// FunctionBlocks/T_SafeMuting
// Model of the TwinSAFE FB MUTING.
// Suppresses the protective device (OSSDIn) while the muting sensors are actuated in the expected order.
// Sequence (sequential inputs, four sensors, forward):
//   M1 on, M2 on, OSSD blocked, M3 on, M1 off, M4 on, M2 off, OSSD clear, M3 off, M4 off
// Sequence (two sensors: parallel inputs, or sequential with MutingIn3/4 unconnected):
//   S1 on, S2 on, OSSD blocked, S1 off, OSSD clear, S2 off
// Any other change of a sensor or the OSSD during a sequence violates it (diagnostic bit 6).
// The Safety Editor refuses an EDM reset time that is not 0 ms, a multiple of 10 ms and at most 60000 ms:
// the model then reports Error with diagnostic bit 15 instead of running (see T_SafeFunctionBlockBase).
{attribute 'reflection'}
FUNCTION_BLOCK T_SafeMuting EXTENDS T_SafeFunctionBlockBase
VAR_INPUT
    MutingEnable : BOOL; // may be a standard PLC signal
    EDM1 : BOOL; // feedback loop of MuteOut
    EDM2 : BOOL; // feedback loop of MuteDelOut
    MutingIn1 : BOOL;
    MutingIn2 : BOOL;
    OSSDIn1 : BOOL; // protective device channel 1 (TRUE = clear)
    OSSDIn2 : BOOL; // protective device channel 2
    MutingIn3 : BOOL;
    MutingIn4 : BOOL;
    Parameters : ST_SafeMutingParameters;
END_VAR
VAR_OUTPUT
    MutingActive : BOOL; // muting lamp
    MuteOut : BOOL;
    MuteDelOut : BOOL;
END_VAR
VAR
    {attribute 'is_connected' := 'MutingEnable'}
    _mutingEnableConnected : BOOL;
    {attribute 'is_connected' := 'EDM1'}
    _eDM1Connected : BOOL;
    {attribute 'is_connected' := 'EDM2'}
    _eDM2Connected : BOOL;
    {attribute 'is_connected' := 'MutingIn1'}
    _mutingIn1Connected : BOOL;
    {attribute 'is_connected' := 'MutingIn2'}
    _mutingIn2Connected : BOOL;
    {attribute 'is_connected' := 'OSSDIn1'}
    _oSSDIn1Connected : BOOL;
    {attribute 'is_connected' := 'OSSDIn2'}
    _oSSDIn2Connected : BOOL;
    {attribute 'is_connected' := 'MutingIn3'}
    _mutingIn3Connected : BOOL;
    {attribute 'is_connected' := 'MutingIn4'}
    _mutingIn4Connected : BOOL;
    _pairs : ARRAY[1..3] OF T_SafeInputPair; // 1: MutingIn1/2, 2: MutingIn3/4, 3: OSSDIn1/2
    _state : E_SafeMutingState := E_SafeMutingState.Stop;
    _prevState : E_SafeMutingState;
    _filterTimers : ARRAY[1..4] OF TON;
    _filtered : ARRAY[1..4] OF BOOL;
    _sensor : ARRAY[1..4] OF BOOL; // actuated sensors after configuration
    _ossdBlocked : BOOL;
    _sensorCount : USINT;
    _seqSensor : ARRAY[1..10] OF USINT; // 0 = OSSD
    _seqLevel : ARRAY[1..10] OF BOOL;
    _seqLength : USINT;
    _seqIndex : USINT; // consumed events
    _expected : ARRAY[0..4] OF BOOL; // expected level of each signal (0 = OSSD blocked)
    _maxTimer : TON;
    _delayTimer : TON;
    _pendingError : BOOL;
    _edmResetTimer1 : TON;
    _edmResetTimer2 : TON;
    _edm1Dropped : BOOL;
    _edm2Dropped : BOOL;
END_VAR

SUPER^();

METHOD PRIVATE Actual : BOOL
VAR_INPUT
    signal : USINT; // 0 = OSSD blocked, 1..4 = sensor actuated
END_VAR
IF signal = 0 THEN
    Actual := _ossdBlocked;
ELSE
    Actual := _sensor[signal];
END_IF
END_METHOD

METHOD PRIVATE AddEvent
VAR_INPUT
    sensor : USINT; // 0 = OSSD
    level : BOOL; // sensor actuated / OSSD blocked
    backwards : BOOL;
END_VAR
IF sensor = 0 AND Parameters.OssdCheckOptional THEN
    RETURN;
END_IF

IF _seqLength >= 10 THEN
    RETURN;
END_IF

_seqLength := _seqLength + 1;

IF sensor > 0 AND backwards THEN
    _seqSensor[_seqLength] := _sensorCount + 1 - sensor;
ELSE
    _seqSensor[_seqLength] := sensor;
END_IF

_seqLevel[_seqLength] := level;
END_METHOD

// Consumes every expected event that has occurred, then checks that no signal deviates
// from the expected pattern. Returns TRUE when the sequence has been violated.
METHOD PRIVATE Advance : BOOL
VAR
    progressed : BOOL;
    next : USINT;
    k : USINT;
END_VAR
REPEAT
    progressed := FALSE;

    IF _seqIndex < _seqLength THEN
        next := _seqIndex + 1;

        IF Actual(_seqSensor[next]) = _seqLevel[next] THEN
            _expected[_seqSensor[next]] := _seqLevel[next];
            _seqIndex                   := next;
            progressed                  := TRUE;
        END_IF
    END_IF
UNTIL NOT progressed
END_REPEAT

FOR k := 0 TO _sensorCount DO
    IF k = 0 AND Parameters.OssdCheckOptional THEN
        CONTINUE;
    END_IF

    IF Actual(k) <> _expected[k] THEN
        Advance := TRUE;
    END_IF
END_FOR
END_METHOD

METHOD PRIVATE AnySensor : BOOL
VAR
    k : USINT;
END_VAR
FOR k := 1 TO _sensorCount DO
    AnySensor := AnySensor OR _sensor[k];
END_FOR
END_METHOD

// Builds the expected event list for the configured sensor arrangement.
METHOD PRIVATE BuildSequence
VAR_INPUT
    backwards : BOOL;
END_VAR
_seqLength := 0;

IF _sensorCount = 4 THEN
    AddEvent(1, TRUE, backwards);
    AddEvent(2, TRUE, backwards);
    AddEvent(0, TRUE, backwards);
    AddEvent(3, TRUE, backwards);
    AddEvent(1, FALSE, backwards);
    AddEvent(4, TRUE, backwards);
    AddEvent(2, FALSE, backwards);
    AddEvent(0, FALSE, backwards);
    AddEvent(3, FALSE, backwards);
    AddEvent(4, FALSE, backwards);
ELSE
    AddEvent(1, TRUE, backwards);
    AddEvent(2, TRUE, backwards);
    AddEvent(0, TRUE, backwards);
    AddEvent(1, FALSE, backwards);
    AddEvent(0, FALSE, backwards);
    AddEvent(2, FALSE, backwards);
END_IF
END_METHOD

// The EDM reset times must be 0 ms or a multiple of 10 ms up to 60000 ms (Safety Editor: "'Reset Time' parameter ... has to be 0 ms or a multiple of 10 ms and maximal 60000 ms").
METHOD PROTECTED ConfigurationOk : BOOL
IF NOT F_SafeResetTimeOk(Parameters.Edm1ResetTime) THEN
    _configurationFault := 'T_SafeMuting: $'Reset Time$' parameter of EDM1 of MUTING has to be 0 ms or a multiple of 10 ms and maximal 60000 ms';
    RETURN;
ELSIF NOT F_SafeResetTimeOk(Parameters.Edm2ResetTime) THEN
    _configurationFault := 'T_SafeMuting: $'Reset Time$' parameter of EDM2 of MUTING has to be 0 ms or a multiple of 10 ms and maximal 60000 ms';
    RETURN;
END_IF

ConfigurationOk := TRUE;
END_METHOD

// Checks the EDM inputs at restart and records diagnostic bits 4/5 on failure.
METHOD PRIVATE EdmInputsOk : BOOL
EdmInputsOk := TRUE;

IF _eDM1Connected AND NOT EDM1 THEN
    SetDiagBit(4);
    EdmInputsOk := FALSE;
END_IF

IF _eDM2Connected AND NOT EDM2 THEN
    SetDiagBit(5);
    EdmInputsOk := FALSE;
END_IF
END_METHOD

// TRUE when every connected EDM input reads 1 (contactors released).
METHOD PRIVATE EdmInputsTrue : BOOL
EdmInputsTrue := (NOT _eDM1Connected OR EDM1) AND (NOT _eDM2Connected OR EDM2);
END_METHOD

// EL6910 extension: after the outputs switch on, each connected EDM input must drop to FALSE
// within its Reset Time. Returns FALSE (and sets diagnostic bits 4/5) on timeout.
METHOD PRIVATE EdmResetOk : BOOL
EdmResetOk := TRUE;

IF _eDM1Connected AND Parameters.Edm1ResetTime > T#0S THEN
    IF NOT EDM1 THEN
        _edm1Dropped := TRUE;
    END_IF

    _edmResetTimer1(IN := NOT _edm1Dropped, PT := Parameters.Edm1ResetTime);

    IF _edmResetTimer1.Q THEN
        SetDiagBit(4);
        EdmResetOk := FALSE;
    END_IF
END_IF

IF _eDM2Connected AND Parameters.Edm2ResetTime > T#0S THEN
    IF NOT EDM2 THEN
        _edm2Dropped := TRUE;
    END_IF

    _edmResetTimer2(IN := NOT _edm2Dropped, PT := Parameters.Edm2ResetTime);

    IF _edmResetTimer2.Q THEN
        SetDiagBit(5);
        EdmResetOk := FALSE;
    END_IF
END_IF
END_METHOD

METHOD PRIVATE IsMuting : BOOL
IsMuting := (TO_BYTE(_state) >= TO_BYTE(E_SafeMutingState.Muting1)) AND (TO_BYTE(_state) <= TO_BYTE(E_SafeMutingState.Muting9));
END_METHOD

PROPERTY MutingState : E_SafeMutingState
GET
MutingState := _state;
END_GET
END_PROPERTY

// State code for the given number of consumed sequence events.
METHOD PRIVATE MutingStateFor : E_SafeMutingState
VAR_INPUT
    consumed : USINT;
END_VAR
CASE consumed OF
    1:
        MutingStateFor := E_SafeMutingState.Muting1;
    2:
        MutingStateFor := E_SafeMutingState.Muting2;
    3:
        MutingStateFor := E_SafeMutingState.Muting3;
    4:
        MutingStateFor := E_SafeMutingState.Muting4;
    5:
        MutingStateFor := E_SafeMutingState.Muting5;
    6:
        MutingStateFor := E_SafeMutingState.Muting6;
    7:
        MutingStateFor := E_SafeMutingState.Muting7;
    8:
        MutingStateFor := E_SafeMutingState.Muting8;
    9:
        MutingStateFor := E_SafeMutingState.Muting9;
ELSE
    MutingStateFor := E_SafeMutingState.Run;
END_CASE
END_METHOD

METHOD PROTECTED Process
VAR
    raw : ARRAY[1..4] OF BOOL;
    i : USINT;
    acknowledge : BOOL;
    discError : BOOL;
    operating : BOOL;
    startFwd : BOOL;
    startBwd : BOOL;
    k : USINT;
    stateBefore : E_SafeMutingState;
    passes : USINT;
END_VAR
// Debounce of the muting inputs
raw[1] := MutingIn1;
raw[2] := MutingIn2;
raw[3] := MutingIn3;
raw[4] := MutingIn4;

FOR i := 1 TO 4 DO
    _filterTimers[i](IN := (raw[i] <> _filtered[i]), PT := Parameters.FilterTime);

    IF _filterTimers[i].Q OR Parameters.FilterTime = T#0S THEN
        _filtered[i] := raw[i];
    END_IF
END_FOR

acknowledge := (_state = E_SafeMutingState.Error) AND _errAck;
_pairs[1](
    In1 := _filtered[1],
    In2 := _filtered[2],
    Active1 := _mutingIn1Connected,
    Active2 := _mutingIn2Connected,
    MakeContact1 := Parameters.MutingIn1MakeContact,
    MakeContact2 := Parameters.MutingIn2MakeContact,
    DiscrepancyTime := Parameters.MutingDiscrepancyTime1,
    Monitor := _fbRun AND NOT Parameters.SequentialInputs,
    SafeInputsAfterDiscError := Parameters.SafeInputsAfterDiscError,
    Acknowledge := acknowledge
);

_pairs[2](
    In1 := _filtered[3],
    In2 := _filtered[4],
    Active1 := _mutingIn3Connected,
    Active2 := _mutingIn4Connected,
    MakeContact1 := Parameters.MutingIn3MakeContact,
    MakeContact2 := Parameters.MutingIn4MakeContact,
    DiscrepancyTime := Parameters.MutingDiscrepancyTime2,
    Monitor := _fbRun AND NOT Parameters.SequentialInputs,
    SafeInputsAfterDiscError := Parameters.SafeInputsAfterDiscError,
    Acknowledge := acknowledge
);

_pairs[3](
    In1 := OSSDIn1,
    In2 := OSSDIn2,
    Active1 := _oSSDIn1Connected,
    Active2 := _oSSDIn2Connected,
    MakeContact1 := Parameters.OSSDIn1MakeContact,
    MakeContact2 := Parameters.OSSDIn2MakeContact,
    DiscrepancyTime := Parameters.OssdDiscrepancyTime,
    Monitor := _fbRun,
    SafeInputsAfterDiscError := Parameters.SafeInputsAfterDiscError,
    Acknowledge := acknowledge
);

IF Parameters.SequentialInputs THEN
    _sensorCount := SEL(_mutingIn3Connected OR _mutingIn4Connected, 2, 4);
    _sensor[1]   := F_SafeInputValue(_mutingIn1Connected, Parameters.MutingIn1MakeContact, _filtered[1]);
    _sensor[2]   := F_SafeInputValue(_mutingIn2Connected, Parameters.MutingIn2MakeContact, _filtered[2]);
    _sensor[3]   := F_SafeInputValue(_mutingIn3Connected, Parameters.MutingIn3MakeContact, _filtered[3]);
    _sensor[4]   := F_SafeInputValue(_mutingIn4Connected, Parameters.MutingIn4MakeContact, _filtered[4]);
ELSE
    _sensorCount := 2;
    _sensor[1]   := _pairs[1].IsActive AND _pairs[1].AllTrue;
    _sensor[2]   := _pairs[2].IsActive AND _pairs[2].AllTrue;
    _sensor[3]   := FALSE;
    _sensor[4]   := FALSE;
END_IF

_ossdBlocked := NOT _pairs[3].AllTrue;

FOR i := 1 TO 3 DO
    discError := discError OR _pairs[i].DiscrepancyError;
END_FOR

IF NOT _fbRun AND _state <> E_SafeMutingState.Error AND _state <> E_SafeMutingState.Reset THEN
    _state := E_SafeMutingState.Stop;
END_IF

operating := (_state = E_SafeMutingState.Safe) OR (_state = E_SafeMutingState.Run) OR IsMuting();

IF discError THEN
    IF operating THEN
        UpdateDiscrepancyDiag();
        _state := E_SafeMutingState.Error;
    ELSIF _state = E_SafeMutingState.DelayOut THEN
        UpdateDiscrepancyDiag();
        _pendingError := TRUE;
    END_IF
END_IF

passes := 0;

REPEAT
    stateBefore := _state;

    CASE _state OF
        E_SafeMutingState.Stop:
            IF StateChanged() THEN
                SetOutputsSafe();
                MutingActive  := FALSE;
                Error         := FALSE;
                Diag          := 0;
                _pendingError := FALSE;
            END_IF

            IF _fbRun THEN
                _state := E_SafeMutingState.Safe;
            END_IF

        E_SafeMutingState.Safe:
            IF StateChanged() THEN
                SetOutputsSafe();
                MutingActive := FALSE;
            END_IF

            IF NOT _ossdBlocked AND EdmInputsTrue() THEN
                _state := E_SafeMutingState.Run;
            END_IF

        E_SafeMutingState.Run:
            IF StateChanged() THEN
                MuteOut      := TRUE;
                MuteDelOut   := TRUE;
                MutingActive := FALSE;
                StartEdmResetMonitoring();
                _seqIndex := 0;
                _maxTimer(IN := FALSE, PT := Parameters.MaxMutingTime);
            END_IF

            startFwd := _sensor[1];
            startBwd := Parameters.BackwardsMode AND _sensor[_sensorCount];

            IF NOT EdmResetOk() THEN
                _state := E_SafeMutingState.Error;
            ELSIF MutingEnable AND (startFwd OR startBwd) THEN
                BuildSequence(startBwd AND NOT startFwd);

                FOR k := 0 TO 4 DO
                    _expected[k] := FALSE;
                END_FOR

                _seqIndex := 0;

                IF Advance() THEN
                    SetDiagBit(6);
                    _state := E_SafeMutingState.Error;
                ELSE
                    _state := MutingStateFor(_seqIndex);
                END_IF
            ELSIF MutingEnable AND AnySensor() THEN
                // a sensor actuated out of order while muting is enabled violates the sequence
                SetDiagBit(6);
                _state := E_SafeMutingState.Error;
            ELSIF _ossdBlocked THEN
                IF Parameters.DelayTime > T#0S THEN
                    _state := E_SafeMutingState.DelayOut;
                ELSE
                    _state := E_SafeMutingState.Safe;
                END_IF
            END_IF

        E_SafeMutingState.Muting1,
        E_SafeMutingState.Muting2,
        E_SafeMutingState.Muting3,
        E_SafeMutingState.Muting4,
        E_SafeMutingState.Muting5,
        E_SafeMutingState.Muting6,
        E_SafeMutingState.Muting7,
        E_SafeMutingState.Muting8,
        E_SafeMutingState.Muting9:
            IF StateChanged() THEN
                MuteOut      := TRUE;
                MuteDelOut   := TRUE;
                MutingActive := TRUE;
            END_IF

            _maxTimer(IN := (Parameters.MaxMutingTime > T#0S), PT := Parameters.MaxMutingTime);

            IF NOT MutingEnable THEN
                // muting withdrawn: the protective device takes over immediately
                IF NOT _ossdBlocked THEN
                    _state := E_SafeMutingState.Run;
                ELSIF Parameters.DelayTime > T#0S THEN
                    _state := E_SafeMutingState.DelayOut;
                ELSE
                    _state := E_SafeMutingState.Safe;
                END_IF
            ELSIF _maxTimer.Q THEN
                SetDiagBit(7);
                _state := E_SafeMutingState.Error;
            ELSIF Advance() THEN
                SetDiagBit(6);
                _state := E_SafeMutingState.Error;
            ELSIF _seqIndex >= _seqLength THEN
                _state := E_SafeMutingState.Run;
            ELSE
                _state := MutingStateFor(_seqIndex);
            END_IF

        E_SafeMutingState.DelayOut:
            IF StateChanged() THEN
                MuteOut      := FALSE;
                MuteDelOut   := TRUE;
                MutingActive := FALSE;
                _delayTimer(IN := FALSE, PT := Parameters.DelayTime);
            END_IF

            _delayTimer(IN := TRUE, PT := Parameters.DelayTime);

            IF _delayTimer.Q THEN
                _state := SEL(_pendingError, E_SafeMutingState.Safe, E_SafeMutingState.Error);
            END_IF

        E_SafeMutingState.Error:
            IF StateChanged() THEN
                SetOutputsSafe();
                MutingActive  := FALSE;
                Error         := TRUE;
                _pendingError := FALSE;
            END_IF

            UpdateDiscrepancyDiag();

            IF _errAck AND NOT discError THEN
                _state := E_SafeMutingState.Reset;
            END_IF

        E_SafeMutingState.Reset:
            IF StateChanged() THEN
                SetOutputsSafe();
                Error := FALSE;
                Diag  := 0;
            END_IF

            IF _errAckFallingEdge THEN
                _state := SEL(_fbRun, E_SafeMutingState.Stop, E_SafeMutingState.Safe);
            END_IF
    END_CASE

    passes := passes + 1;
UNTIL (stateBefore = _state) OR (passes >= 3)
END_REPEAT

State := TO_BYTE(_state);
END_METHOD

METHOD PRIVATE SetOutputsSafe
MuteOut    := FALSE;
MuteDelOut := FALSE;
END_METHOD

METHOD PRIVATE StartEdmResetMonitoring
_edm1Dropped := FALSE;
_edm2Dropped := FALSE;
_edmResetTimer1(IN := FALSE, PT := Parameters.Edm1ResetTime);
_edmResetTimer2(IN := FALSE, PT := Parameters.Edm2ResetTime);
END_METHOD

METHOD PRIVATE StateChanged : BOOL
IF _prevState = _state THEN
    RETURN;
END_IF

_prevState   := _state;
StateChanged := TRUE;
END_METHOD

// Mirrors the discrepancy state of every pair into the diagnostic bits.
METHOD PRIVATE UpdateDiscrepancyDiag
VAR
    i : USINT;
END_VAR
FOR i := 1 TO 3 DO
    IF _pairs[i].DiscrepancyError THEN
        SetDiagBit(SEL(i = 1, SEL(i = 2, 1, 2), 0));

        IF _pairs[i].AwaitingSafeInputs THEN
            SetDiagBit(SEL(i = 1, SEL(i = 2, 9, 10), 8));
        ELSE
            ClearDiagBit(SEL(i = 1, SEL(i = 2, 9, 10), 8));
        END_IF
    END_IF
END_FOR
END_METHOD

END_FUNCTION_BLOCK

// FunctionBlocks/T_SafeOpMode
// Model of the TwinSAFE FB OPMODE (operating mode selector).
// Exactly one connected OpIn input must be TRUE for the matching OpOut to be set.
// Manual restart is active when the Restart port is connected.
// The Safety Editor refuses an OPMODE with fewer than two OpIn ports connected: the model then reports
// Error with diagnostic bit 15 instead of running (see T_SafeFunctionBlockBase).
{attribute 'reflection'}
FUNCTION_BLOCK T_SafeOpMode EXTENDS T_SafeFunctionBlockBase
VAR_INPUT
    Restart : BOOL; // may be a standard PLC signal
    OpIn1 : BOOL;
    OpIn2 : BOOL;
    OpIn3 : BOOL;
    OpIn4 : BOOL;
    OpIn5 : BOOL;
    OpIn6 : BOOL;
    OpIn7 : BOOL;
    OpIn8 : BOOL;
    Parameters : ST_SafeOpModeParameters;
END_VAR
VAR_OUTPUT
    OpOut1 : BOOL;
    OpOut2 : BOOL;
    OpOut3 : BOOL;
    OpOut4 : BOOL;
    OpOut5 : BOOL;
    OpOut6 : BOOL;
    OpOut7 : BOOL;
    OpOut8 : BOOL;
END_VAR
VAR
    {attribute 'is_connected' := 'Restart'}
    _restartConnected : BOOL;
    {attribute 'is_connected' := 'OpIn1'}
    _opIn1Connected : BOOL;
    {attribute 'is_connected' := 'OpIn2'}
    _opIn2Connected : BOOL;
    {attribute 'is_connected' := 'OpIn3'}
    _opIn3Connected : BOOL;
    {attribute 'is_connected' := 'OpIn4'}
    _opIn4Connected : BOOL;
    {attribute 'is_connected' := 'OpIn5'}
    _opIn5Connected : BOOL;
    {attribute 'is_connected' := 'OpIn6'}
    _opIn6Connected : BOOL;
    {attribute 'is_connected' := 'OpIn7'}
    _opIn7Connected : BOOL;
    {attribute 'is_connected' := 'OpIn8'}
    _opIn8Connected : BOOL;
    _state : E_SafeFbState := E_SafeFbState.Stop;
    _prevState : E_SafeFbState;
    _restartPrev : BOOL;
    _discrepancyTimer : TON;
    _modeSelectedBefore : BOOL;
END_VAR

SUPER^();

// At least two OpIn ports must be connected (Safety Editor: "OPMODE does not have at least 2 input ports connected").
METHOD PROTECTED ConfigurationOk : BOOL
VAR
    connectedInputs : USINT;
END_VAR
connectedInputs := BOOL_TO_USINT(_opIn1Connected)
    + BOOL_TO_USINT(_opIn2Connected)
    + BOOL_TO_USINT(_opIn3Connected)
    + BOOL_TO_USINT(_opIn4Connected)
    + BOOL_TO_USINT(_opIn5Connected)
    + BOOL_TO_USINT(_opIn6Connected)
    + BOOL_TO_USINT(_opIn7Connected)
    + BOOL_TO_USINT(_opIn8Connected);

IF connectedInputs < 2 THEN
    _configurationFault := 'T_SafeOpMode: OPMODE does not have at least 2 input ports connected';
    RETURN;
END_IF

ConfigurationOk := TRUE;
END_METHOD

METHOD PROTECTED Process
VAR
    count : USINT;
    selected : USINT;
    exactlyOne : BOOL;
    restartFalling : BOOL;
    monitoring : BOOL;
    operating : BOOL;
    stateBefore : E_SafeFbState;
    passes : USINT;
END_VAR
IF _opIn1Connected AND OpIn1 THEN
    count    := count + 1;
    selected := 1;
END_IF

IF _opIn2Connected AND OpIn2 THEN
    count    := count + 1;
    selected := 2;
END_IF

IF _opIn3Connected AND OpIn3 THEN
    count    := count + 1;
    selected := 3;
END_IF

IF _opIn4Connected AND OpIn4 THEN
    count    := count + 1;
    selected := 4;
END_IF

IF _opIn5Connected AND OpIn5 THEN
    count    := count + 1;
    selected := 5;
END_IF

IF _opIn6Connected AND OpIn6 THEN
    count    := count + 1;
    selected := 6;
END_IF

IF _opIn7Connected AND OpIn7 THEN
    count    := count + 1;
    selected := 7;
END_IF

IF _opIn8Connected AND OpIn8 THEN
    count    := count + 1;
    selected := 8;
END_IF

exactlyOne     := (count = 1);
restartFalling := NOT Restart AND _restartPrev;
_restartPrev   := Restart;

IF NOT _fbRun AND _state <> E_SafeFbState.Error AND _state <> E_SafeFbState.Reset THEN
    _state := E_SafeFbState.Stop;
END_IF

// Discrepancy monitoring of a mode change: none or several inputs set for too long
operating  := (_state = E_SafeFbState.Safe) OR (_state = E_SafeFbState.Start) OR (_state = E_SafeFbState.Run);
monitoring := operating AND _modeSelectedBefore AND NOT exactlyOne AND (Parameters.DiscrepancyTime > T#0S);
_discrepancyTimer(IN := monitoring, PT := Parameters.DiscrepancyTime);

IF _discrepancyTimer.Q AND operating THEN
    SetDiagBit(0);
    _state := E_SafeFbState.Error;
END_IF

passes := 0;

REPEAT
    stateBefore := _state;

    CASE _state OF
        E_SafeFbState.Stop:
            IF StateChanged() THEN
                SetOutputs(0);
                Error               := FALSE;
                Diag                := 0;
                _modeSelectedBefore := FALSE;
            END_IF

            IF _fbRun THEN
                _state := E_SafeFbState.Safe;
            END_IF

        E_SafeFbState.Safe:
            IF StateChanged() THEN
                SetOutputs(0);
            END_IF

            IF exactlyOne THEN
                IF NOT _restartConnected THEN
                    _state := E_SafeFbState.Run;
                ELSIF Restart THEN
                    _state := E_SafeFbState.Start;
                END_IF
            END_IF

        E_SafeFbState.Start:
            IF StateChanged() THEN
                SetOutputs(0);
            END_IF

            IF NOT exactlyOne THEN
                _state := E_SafeFbState.Safe;
            ELSIF restartFalling THEN
                _state := E_SafeFbState.Run;
            END_IF

        E_SafeFbState.Run:
            IF StateChanged() THEN
                _modeSelectedBefore := TRUE;
            END_IF

            IF exactlyOne THEN
                SetOutputs(selected);
            ELSE
                SetOutputs(0);
                _state := E_SafeFbState.Safe;
            END_IF

        E_SafeFbState.Error:
            IF StateChanged() THEN
                SetOutputs(0);
                Error := TRUE;
            END_IF

            IF _errAck THEN
                _state := E_SafeFbState.Reset;
            END_IF

        E_SafeFbState.Reset:
            IF StateChanged() THEN
                Error := FALSE;
                Diag  := 0;
            END_IF

            IF _errAckFallingEdge THEN
                _state := SEL(_fbRun, E_SafeFbState.Stop, E_SafeFbState.Safe);
            END_IF
    END_CASE

    passes := passes + 1;
UNTIL (stateBefore = _state) OR (passes >= 3)
END_REPEAT

State := TO_BYTE(_state);
END_METHOD

METHOD PRIVATE SetOutputs
VAR_INPUT
    selected : USINT; // 0 = all outputs off
END_VAR
OpOut1 := (selected = 1);
OpOut2 := (selected = 2);
OpOut3 := (selected = 3);
OpOut4 := (selected = 4);
OpOut5 := (selected = 5);
OpOut6 := (selected = 6);
OpOut7 := (selected = 7);
OpOut8 := (selected = 8);
END_METHOD

METHOD PRIVATE StateChanged : BOOL
IF _prevState = _state THEN
    RETURN;
END_IF

_prevState   := _state;
StateChanged := TRUE;
END_METHOD

END_FUNCTION_BLOCK

// FunctionBlocks/T_SafeOr
// Model of the TwinSAFE FB OR. Connected inputs are active.
// The Safety Editor refuses an OR with fewer than two OrIn ports connected: the model then reports
// Error with diagnostic bit 15 instead of running (see T_SafeFunctionBlockBase).
{attribute 'reflection'}
FUNCTION_BLOCK T_SafeOr EXTENDS T_SafeFunctionBlockBase
VAR_INPUT
    OrIn1 : BOOL;
    OrIn2 : BOOL;
    OrIn3 : BOOL;
    OrIn4 : BOOL;
    OrIn5 : BOOL;
    OrIn6 : BOOL;
    OrIn7 : BOOL;
    OrIn8 : BOOL;
    Parameters : ST_SafeLogicParameters;
END_VAR
VAR_OUTPUT
    OrOut : BOOL;
END_VAR
VAR
    {attribute 'is_connected' := 'OrIn1'}
    _orIn1Connected : BOOL;
    {attribute 'is_connected' := 'OrIn2'}
    _orIn2Connected : BOOL;
    {attribute 'is_connected' := 'OrIn3'}
    _orIn3Connected : BOOL;
    {attribute 'is_connected' := 'OrIn4'}
    _orIn4Connected : BOOL;
    {attribute 'is_connected' := 'OrIn5'}
    _orIn5Connected : BOOL;
    {attribute 'is_connected' := 'OrIn6'}
    _orIn6Connected : BOOL;
    {attribute 'is_connected' := 'OrIn7'}
    _orIn7Connected : BOOL;
    {attribute 'is_connected' := 'OrIn8'}
    _orIn8Connected : BOOL;
    _state : E_SafeFbState := E_SafeFbState.Stop;
END_VAR

SUPER^();

// At least two OrIn ports must be connected (Safety Editor: "OR does not have at least 2 input ports active and connected").
METHOD PROTECTED ConfigurationOk : BOOL
VAR
    connectedInputs : USINT;
END_VAR
connectedInputs := BOOL_TO_USINT(_orIn1Connected)
    + BOOL_TO_USINT(_orIn2Connected)
    + BOOL_TO_USINT(_orIn3Connected)
    + BOOL_TO_USINT(_orIn4Connected)
    + BOOL_TO_USINT(_orIn5Connected)
    + BOOL_TO_USINT(_orIn6Connected)
    + BOOL_TO_USINT(_orIn7Connected)
    + BOOL_TO_USINT(_orIn8Connected);

IF connectedInputs < 2 THEN
    _configurationFault := 'T_SafeOr: OR does not have at least 2 input ports active and connected';
    RETURN;
END_IF

ConfigurationOk := TRUE;
END_METHOD

METHOD PROTECTED Process
VAR
    result : BOOL;
END_VAR
result := FALSE;
result := result OR F_SafeInputValue(_orIn1Connected, Parameters.In1MakeContact, OrIn1);
result := result OR F_SafeInputValue(_orIn2Connected, Parameters.In2MakeContact, OrIn2);
result := result OR F_SafeInputValue(_orIn3Connected, Parameters.In3MakeContact, OrIn3);
result := result OR F_SafeInputValue(_orIn4Connected, Parameters.In4MakeContact, OrIn4);
result := result OR F_SafeInputValue(_orIn5Connected, Parameters.In5MakeContact, OrIn5);
result := result OR F_SafeInputValue(_orIn6Connected, Parameters.In6MakeContact, OrIn6);
result := result OR F_SafeInputValue(_orIn7Connected, Parameters.In7MakeContact, OrIn7);
result := result OR F_SafeInputValue(_orIn8Connected, Parameters.In8MakeContact, OrIn8);

IF NOT _fbRun THEN
    _state := E_SafeFbState.Stop;
ELSIF result THEN
    _state := E_SafeFbState.Run;
ELSE
    _state := E_SafeFbState.Safe;
END_IF

OrOut := (_state = E_SafeFbState.Run);
Error := FALSE;
Diag  := 0;
State := TO_BYTE(_state);
END_METHOD

END_FUNCTION_BLOCK

// FunctionBlocks/T_SafeSr
// Model of the TwinSAFE FB SR (set dominant latch).
// The Safety Editor refuses an SR with Set or Reset unconnected: the model then reports Error with
// diagnostic bit 15 instead of running (see T_SafeFunctionBlockBase).
{attribute 'reflection'}
FUNCTION_BLOCK T_SafeSr EXTENDS T_SafeFunctionBlockBase
VAR_INPUT
    Set : BOOL;
    Reset : BOOL;
    Parameters : ST_SafeLatchParameters;
END_VAR
VAR_OUTPUT
    SrOut : BOOL;
END_VAR
VAR
    {attribute 'is_connected' := 'Set'}
    _setConnected : BOOL;
    {attribute 'is_connected' := 'Reset'}
    _resetConnected : BOOL;
    _state : E_SafeLatchState := E_SafeLatchState.Stop;
END_VAR

SUPER^();

// Set and Reset must both be connected (Safety Editor: "Inport Set of SR must be connected").
METHOD PROTECTED ConfigurationOk : BOOL
IF NOT _setConnected THEN
    _configurationFault := 'T_SafeSr: Inport Set of SR must be connected';
    RETURN;
ELSIF NOT _resetConnected THEN
    _configurationFault := 'T_SafeSr: Inport Reset of SR must be connected';
    RETURN;
END_IF

ConfigurationOk := TRUE;
END_METHOD

METHOD PROTECTED Process
VAR
    setActive : BOOL;
    resetActive : BOOL;
END_VAR
setActive   := F_SafeInputValue(_setConnected, Parameters.SetMakeContact, Set);
resetActive := F_SafeInputValue(_resetConnected, Parameters.ResetMakeContact, Reset);

IF NOT _fbRun THEN
    _state := E_SafeLatchState.Stop;
ELSE
    IF _state = E_SafeLatchState.Stop THEN
        _state := E_SafeLatchState.Safe;
    END_IF

    IF setActive THEN
        _state := E_SafeLatchState.Set;
    ELSIF resetActive THEN
        _state := E_SafeLatchState.Safe;
    END_IF
END_IF

SrOut := (_state = E_SafeLatchState.Set);
Error := FALSE;
Diag  := 0;
State := TO_BYTE(_state);
END_METHOD

END_FUNCTION_BLOCK

// FunctionBlocks/T_SafeTof
// Model of the TwinSAFE FB TOF (switch-off delay).
// The Safety Editor refuses a TOF with TofIn1 unconnected: the model then reports Error with diagnostic
// bit 15 instead of running (see T_SafeFunctionBlockBase).
{attribute 'reflection'}
FUNCTION_BLOCK T_SafeTof EXTENDS T_SafeFunctionBlockBase
VAR_INPUT
    TofIn1 : BOOL;
    Parameters : ST_SafeTimerParameters;
END_VAR
VAR_OUTPUT
    TofOut : BOOL;
END_VAR
VAR
    {attribute 'is_connected' := 'TofIn1'}
    _tofIn1Connected : BOOL;
    _state : E_SafeFbState := E_SafeFbState.Stop;
    _timer : TOF;
END_VAR

SUPER^();

// TofIn1 must be connected (Safety Editor: "Inport TofIn1 of TOF must be connected").
METHOD PROTECTED ConfigurationOk : BOOL
IF NOT _tofIn1Connected THEN
    _configurationFault := 'T_SafeTof: Inport TofIn1 of TOF must be connected';
    RETURN;
END_IF

ConfigurationOk := TRUE;
END_METHOD

METHOD PROTECTED Process
VAR
    inputActive : BOOL;
END_VAR
inputActive := F_SafeInputValue(_tofIn1Connected, Parameters.MakeContact, TofIn1);

IF NOT _fbRun THEN
    // a stopped FB does not run its delay
    _timer(IN := FALSE, PT := T#0S);
    _state := E_SafeFbState.Stop;
ELSE
    _timer(IN := inputActive, PT := Parameters.DelayTime);

    IF inputActive THEN
        _state := E_SafeFbState.Run;
    ELSIF _timer.Q THEN
        _state := E_SafeFbState.DelayOut;
    ELSE
        _state := E_SafeFbState.Safe;
    END_IF
END_IF

TofOut := (_state = E_SafeFbState.Run) OR (_state = E_SafeFbState.DelayOut);
Error  := FALSE;
Diag   := 0;
State  := TO_BYTE(_state);
END_METHOD

END_FUNCTION_BLOCK

// FunctionBlocks/T_SafeTwoHand
// Model of the TwinSAFE FB TWOHAND (two-hand control).
// Both hands (input pairs) must be actuated, optionally within HandDiscrepancyTime of each other.
// The output can only be set again after both hands were released together.
{attribute 'reflection'}
FUNCTION_BLOCK T_SafeTwoHand EXTENDS T_SafeFunctionBlockBase
VAR_INPUT
    Twohand1 : BOOL; // first hand, channel 1
    Twohand2 : BOOL; // first hand, channel 2
    Twohand3 : BOOL; // second hand, channel 1
    Twohand4 : BOOL; // second hand, channel 2
    Parameters : ST_SafeTwoHandParameters;
END_VAR
VAR_OUTPUT
    TwoHandOut : BOOL;
END_VAR
VAR
    {attribute 'is_connected' := 'Twohand1'}
    _twohand1Connected : BOOL;
    {attribute 'is_connected' := 'Twohand2'}
    _twohand2Connected : BOOL;
    {attribute 'is_connected' := 'Twohand3'}
    _twohand3Connected : BOOL;
    {attribute 'is_connected' := 'Twohand4'}
    _twohand4Connected : BOOL;
    _pairs : ARRAY[1..2] OF T_SafeInputPair;
    _state : E_SafeTwoHandState := E_SafeTwoHandState.Stop;
    _prevState : E_SafeTwoHandState;
    _handTimer : TON;
    _awaitingRelease : BOOL; // between-hands discrepancy error waits for both hands released
END_VAR

SUPER^();

METHOD PROTECTED Process
VAR
    acknowledge : BOOL;
    hand1 : BOOL; // first hand fully actuated
    hand2 : BOOL; // second hand fully actuated
    anyFalse : BOOL; // at least one active input released
    allFalse : BOOL; // every active input released
    discError : BOOL;
    operating : BOOL;
    stateBefore : E_SafeTwoHandState;
    passes : USINT;
END_VAR
acknowledge := (_state = E_SafeTwoHandState.Error) AND _errAck AND NOT _awaitingRelease;
_pairs[1](
    In1 := Twohand1,
    In2 := Twohand2,
    Active1 := _twohand1Connected,
    Active2 := _twohand2Connected,
    MakeContact1 := Parameters.Twohand1MakeContact,
    MakeContact2 := Parameters.Twohand2MakeContact,
    DiscrepancyTime := Parameters.DiscrepancyTime1,
    Monitor := _fbRun,
    SafeInputsAfterDiscError := Parameters.SafeInputsAfterDiscError,
    Acknowledge := acknowledge
);

_pairs[2](
    In1 := Twohand3,
    In2 := Twohand4,
    Active1 := _twohand3Connected,
    Active2 := _twohand4Connected,
    MakeContact1 := Parameters.Twohand3MakeContact,
    MakeContact2 := Parameters.Twohand4MakeContact,
    DiscrepancyTime := Parameters.DiscrepancyTime2,
    Monitor := _fbRun,
    SafeInputsAfterDiscError := Parameters.SafeInputsAfterDiscError,
    Acknowledge := acknowledge
);

hand1     := _pairs[1].IsActive AND _pairs[1].AllTrue;
hand2     := _pairs[2].IsActive AND _pairs[2].AllTrue;
anyFalse  := NOT (_pairs[1].AllTrue AND _pairs[2].AllTrue);
allFalse  := (NOT _pairs[1].IsActive OR _pairs[1].AllFalse) AND (NOT _pairs[2].IsActive OR _pairs[2].AllFalse);
discError := _pairs[1].DiscrepancyError OR _pairs[2].DiscrepancyError;

IF NOT _fbRun AND _state <> E_SafeTwoHandState.Error AND _state <> E_SafeTwoHandState.Reset THEN
    _state := E_SafeTwoHandState.Stop;
END_IF

operating := (_state = E_SafeTwoHandState.Safe)
                 OR (_state = E_SafeTwoHandState.OneButton)
                 OR (_state = E_SafeTwoHandState.TwoButton)
                 OR (_state = E_SafeTwoHandState.Run)
                 OR (_state = E_SafeTwoHandState.Release);

IF discError AND operating THEN
    UpdateDiscrepancyDiag();
    _state := E_SafeTwoHandState.Error;
END_IF

IF _awaitingRelease AND allFalse THEN
    _awaitingRelease := FALSE;
END_IF

passes := 0;

REPEAT
    stateBefore := _state;

    CASE _state OF
        E_SafeTwoHandState.Stop:
            IF StateChanged() THEN
                TwoHandOut := FALSE;
                Error      := FALSE;
                Diag       := 0;
            END_IF

            IF _fbRun THEN
                _state := E_SafeTwoHandState.Safe;
            END_IF

        E_SafeTwoHandState.Safe:
            IF StateChanged() THEN
                TwoHandOut := FALSE;
            END_IF

            IF hand1 THEN
                _state := E_SafeTwoHandState.OneButton;
            ELSIF hand2 THEN
                _state := E_SafeTwoHandState.TwoButton;
            END_IF

        E_SafeTwoHandState.OneButton:
            IF StateChanged() THEN
                _handTimer(IN := FALSE, PT := Parameters.HandDiscrepancyTime);
            END_IF

            _handTimer(IN := (Parameters.HandDiscrepancyTime > T#0S), PT := Parameters.HandDiscrepancyTime);

            IF _handTimer.Q THEN
                SetHandDiscrepancyError();
            ELSIF hand1 AND hand2 THEN
                _state := E_SafeTwoHandState.Run;
            ELSIF hand2 THEN
                // second hand actuated while the first is no longer detected
                SetDiagBit(6);
                _state := E_SafeTwoHandState.Error;
            ELSIF NOT hand1 THEN
                _state := SEL(allFalse, E_SafeTwoHandState.Release, E_SafeTwoHandState.Safe);
            END_IF

        E_SafeTwoHandState.TwoButton:
            IF StateChanged() THEN
                _handTimer(IN := FALSE, PT := Parameters.HandDiscrepancyTime);
            END_IF

            _handTimer(IN := (Parameters.HandDiscrepancyTime > T#0S), PT := Parameters.HandDiscrepancyTime);

            IF _handTimer.Q THEN
                SetHandDiscrepancyError();
            ELSIF hand1 AND hand2 THEN
                _state := E_SafeTwoHandState.Run;
            ELSIF hand1 THEN
                SetDiagBit(6);
                _state := E_SafeTwoHandState.Error;
            ELSIF NOT hand2 THEN
                _state := SEL(allFalse, E_SafeTwoHandState.Release, E_SafeTwoHandState.Safe);
            END_IF

        E_SafeTwoHandState.Run:
            IF StateChanged() THEN
                TwoHandOut := TRUE;
            END_IF

            IF anyFalse THEN
                _state := E_SafeTwoHandState.Release;
            END_IF

        E_SafeTwoHandState.Release:
            IF StateChanged() THEN
                TwoHandOut := FALSE;
            END_IF

            IF allFalse THEN
                _state := E_SafeTwoHandState.Safe;
            END_IF

        E_SafeTwoHandState.Error:
            IF StateChanged() THEN
                TwoHandOut := FALSE;
                Error      := TRUE;
            END_IF

            UpdateDiscrepancyDiag();

            IF _awaitingRelease THEN
                SetDiagBit(10);
            ELSE
                ClearDiagBit(10);
            END_IF

            IF _errAck AND NOT _awaitingRelease AND NOT discError THEN
                _state := E_SafeTwoHandState.Reset;
            END_IF

        E_SafeTwoHandState.Reset:
            IF StateChanged() THEN
                TwoHandOut := FALSE;
                Error      := FALSE;
                Diag       := 0;
            END_IF

            IF _errAckFallingEdge THEN
                _state := SEL(_fbRun, E_SafeTwoHandState.Stop, E_SafeTwoHandState.Safe);
            END_IF
    END_CASE

    passes := passes + 1;
UNTIL (stateBefore = _state) OR (passes >= 3)
END_REPEAT

State := TO_BYTE(_state);
END_METHOD

METHOD PRIVATE SetHandDiscrepancyError
SetDiagBit(2);
_awaitingRelease := Parameters.SafeInputsAfterDiscError;
_state           := E_SafeTwoHandState.Error;
END_METHOD

METHOD PRIVATE StateChanged : BOOL
IF _prevState = _state THEN
    RETURN;
END_IF

_prevState   := _state;
StateChanged := TRUE;
END_METHOD

PROPERTY TwoHandState : E_SafeTwoHandState
GET
TwoHandState := _state;
END_GET
END_PROPERTY

// Mirrors the discrepancy state of every pair into the diagnostic bits.
METHOD PRIVATE UpdateDiscrepancyDiag
VAR
    i : USINT;
END_VAR
FOR i := 1 TO 2 DO
    IF _pairs[i].DiscrepancyError THEN
        SetDiagBit(i - 1);

        IF _pairs[i].AwaitingSafeInputs THEN
            SetDiagBit(i + 7);
        ELSE
            ClearDiagBit(i + 7);
        END_IF
    END_IF
END_FOR
END_METHOD

END_FUNCTION_BLOCK

// FunctionBlocks/T_SafeXor
// Model of the TwinSAFE FB XOR: eight independent exclusive-or pairs. A pair is active when connected.
{attribute 'reflection'}
FUNCTION_BLOCK T_SafeXor EXTENDS T_SafeFunctionBlockBase
VAR_INPUT
    Xor1In1 : BOOL;
    Xor2In1 : BOOL;
    Xor1In2 : BOOL;
    Xor2In2 : BOOL;
    Xor1In3 : BOOL;
    Xor2In3 : BOOL;
    Xor1In4 : BOOL;
    Xor2In4 : BOOL;
    Xor1In5 : BOOL;
    Xor2In5 : BOOL;
    Xor1In6 : BOOL;
    Xor2In6 : BOOL;
    Xor1In7 : BOOL;
    Xor2In7 : BOOL;
    Xor1In8 : BOOL;
    Xor2In8 : BOOL;
END_VAR
VAR_OUTPUT
    XorOut1 : BOOL;
    XorOut2 : BOOL;
    XorOut3 : BOOL;
    XorOut4 : BOOL;
    XorOut5 : BOOL;
    XorOut6 : BOOL;
    XorOut7 : BOOL;
    XorOut8 : BOOL;
END_VAR
VAR
    {attribute 'is_connected' := 'Xor1In1'}
    _xor1In1Connected : BOOL;
    {attribute 'is_connected' := 'Xor1In2'}
    _xor1In2Connected : BOOL;
    {attribute 'is_connected' := 'Xor1In3'}
    _xor1In3Connected : BOOL;
    {attribute 'is_connected' := 'Xor1In4'}
    _xor1In4Connected : BOOL;
    {attribute 'is_connected' := 'Xor1In5'}
    _xor1In5Connected : BOOL;
    {attribute 'is_connected' := 'Xor1In6'}
    _xor1In6Connected : BOOL;
    {attribute 'is_connected' := 'Xor1In7'}
    _xor1In7Connected : BOOL;
    {attribute 'is_connected' := 'Xor1In8'}
    _xor1In8Connected : BOOL;
    {attribute 'is_connected' := 'Xor2In1'}
    _xor2In1Connected : BOOL;
    {attribute 'is_connected' := 'Xor2In2'}
    _xor2In2Connected : BOOL;
    {attribute 'is_connected' := 'Xor2In3'}
    _xor2In3Connected : BOOL;
    {attribute 'is_connected' := 'Xor2In4'}
    _xor2In4Connected : BOOL;
    {attribute 'is_connected' := 'Xor2In5'}
    _xor2In5Connected : BOOL;
    {attribute 'is_connected' := 'Xor2In6'}
    _xor2In6Connected : BOOL;
    {attribute 'is_connected' := 'Xor2In7'}
    _xor2In7Connected : BOOL;
    {attribute 'is_connected' := 'Xor2In8'}
    _xor2In8Connected : BOOL;
    _state : E_SafeFbState := E_SafeFbState.Stop;
END_VAR

SUPER^();

METHOD PROTECTED Process
VAR
    run : BOOL;
END_VAR
run     := _fbRun;
_state  := SEL(run, E_SafeFbState.Stop, E_SafeFbState.Run);
XorOut1 := run AND (_xor1In1Connected OR _xor2In1Connected) AND (Xor1In1 XOR Xor2In1);
XorOut2 := run AND (_xor1In2Connected OR _xor2In2Connected) AND (Xor1In2 XOR Xor2In2);
XorOut3 := run AND (_xor1In3Connected OR _xor2In3Connected) AND (Xor1In3 XOR Xor2In3);
XorOut4 := run AND (_xor1In4Connected OR _xor2In4Connected) AND (Xor1In4 XOR Xor2In4);
XorOut5 := run AND (_xor1In5Connected OR _xor2In5Connected) AND (Xor1In5 XOR Xor2In5);
XorOut6 := run AND (_xor1In6Connected OR _xor2In6Connected) AND (Xor1In6 XOR Xor2In6);
XorOut7 := run AND (_xor1In7Connected OR _xor2In7Connected) AND (Xor1In7 XOR Xor2In7);
XorOut8 := run AND (_xor1In8Connected OR _xor2In8Connected) AND (Xor1In8 XOR Xor2In8);
Error   := FALSE;
Diag    := 0;
State   := TO_BYTE(_state);
END_METHOD

END_FUNCTION_BLOCK

// Project Information/F_GetCompany
// This function has been automatically generated from the project information.
{attribute 'signature_flag' := '1073741824'}
{attribute 'TcGenerated'}
{attribute 'no-analysis'}
FUNCTION F_GetCompany : WSTRING
VAR_INPUT
	
END_VAR

F_GetCompany := "Intecre Ltd";

END_FUNCTION

// Project Information/F_GetTitle
// This function has been automatically generated from the project information.
{attribute 'signature_flag' := '1073741824'}
{attribute 'TcGenerated'}
{attribute 'no-analysis'}
FUNCTION F_GetTitle : WSTRING
VAR_INPUT
	
END_VAR

F_GetTitle := "Intecre.TwinSAFE.Models";

END_FUNCTION

// Project Information/F_GetVersion
// This function has been automatically generated from the project information.
{attribute 'signature_flag' := '1073741824'}
{attribute 'TcGenerated'}
{attribute 'no-analysis'}
FUNCTION F_GetVersion : ST_LibVersion
VAR_INPUT
	
END_VAR

F_GetVersion.iMajor := 0;
F_GetVersion.iMinor := 5;
F_GetVersion.iBuild := 0;
F_GetVersion.iRevision := 3;
F_GetVersion.sVersion := '0.5.0.3';
F_GetVersion.nFlags := 0;

END_FUNCTION

// Tests/User_FB_Tests/T_SafePulse_UserFB_Tests
// Tests of the example user FB T_SafePulse_UserFB: TonOut is a pulse of DelayTime while TonIn1 is held.
FUNCTION_BLOCK T_SafePulse_UserFB_Tests EXTENDS TcUnit.FB_TestSuite
VAR
    // Test_PulseForDelayTimeWhileInputHeld
    group_1 : T_SafeGroup;
    fb_1 : T_SafePulse_UserFB(group := group_1) := (Parameters := (DelayTime := T#100MS));
    state_1 : INT := 10;
    waitTimer_1 : TON;
    // Test_PulseEndsWhenInputDrops
    group_2 : T_SafeGroup;
    fb_2 : T_SafePulse_UserFB(group := group_2) := (Parameters := (DelayTime := T#100MS));
    // Test_StoppedGivesNoOutput
    group_3 : T_SafeGroup;
    fb_3 : T_SafePulse_UserFB(group := group_3) := (Parameters := (DelayTime := T#100MS));
    // Test_InnerBlocksJoinTheGroup
    group_4 : T_SafeGroup;
    fb_4 : T_SafePulse_UserFB(group := group_4);
END_VAR

Test_PulseForDelayTimeWhileInputHeld();
Test_PulseEndsWhenInputDrops();
Test_StoppedGivesNoOutput();
Test_InnerBlocksJoinTheGroup();

METHOD PRIVATE Test_InnerBlocksJoinTheGroup
TcUnit.TEST(__POUNAME());
// assert: the composite registered itself and passed the group on to its TON and AND
AssertEquals_UINT(Expected := 3, Actual := group_4.FunctionBlockCount, Message := 'composite and its two inner blocks registered');
TEST_FINISHED_NAMED(__POUNAME());
END_METHOD

METHOD PRIVATE Test_PulseEndsWhenInputDrops
TcUnit.TEST(__POUNAME());
// act / assert
group_2(Run := TRUE);
fb_2(TonIn1 := TRUE);
AssertEquals_BOOL(Expected := TRUE, Actual := fb_2.TonOut, Message := 'pulse on');
AssertEquals_BOOL(Expected := TRUE, Actual := fb_2.IsRunning, Message := 'reports Run to the group while it runs');
fb_2(TonIn1 := FALSE);
AssertEquals_BOOL(Expected := FALSE, Actual := fb_2.TonOut, Message := 'pulse cut off when the input drops');
TEST_FINISHED_NAMED(__POUNAME());
END_METHOD

METHOD PRIVATE Test_PulseForDelayTimeWhileInputHeld
TcUnit.TEST(__POUNAME());
waitTimer_1();

CASE state_1 OF
    10:
        // act: input on, the pulse starts
        group_1(Run := TRUE);
        fb_1(TonIn1 := TRUE);
        // assert
        AssertEquals_BOOL(Expected := TRUE, Actual := fb_1.TonOut, Message := 'pulse starts with the input');
        state_1 := 20;
        waitTimer_1(IN := TRUE, PT := T#50MS);
    20:
        group_1(Run := TRUE);
        fb_1(TonIn1 := TRUE);

        IF NOT waitTimer_1.Q THEN
            RETURN;
        END_IF

        waitTimer_1(IN := FALSE);
        // assert: still inside the delay time
        AssertEquals_BOOL(Expected := TRUE, Actual := fb_1.TonOut, Message := 'pulse still on inside the delay time');
        state_1 := 30;
        waitTimer_1(IN := TRUE, PT := T#200MS);
    30:
        group_1(Run := TRUE);
        fb_1(TonIn1 := TRUE);

        IF NOT waitTimer_1.Q THEN
            RETURN;
        END_IF

        waitTimer_1(IN := FALSE);
        // assert: the delay has elapsed, the pulse is over although the input is still held
        AssertEquals_BOOL(Expected := FALSE, Actual := fb_1.TonOut, Message := 'pulse ends after the delay time');
        // act: release and re-apply the input
        fb_1(TonIn1 := FALSE);
        AssertEquals_BOOL(Expected := FALSE, Actual := fb_1.TonOut, Message := 'no output with the input off');
        fb_1(TonIn1 := TRUE);
        AssertEquals_BOOL(Expected := TRUE, Actual := fb_1.TonOut, Message := 'a new pulse starts on the next rising edge');
        TEST_FINISHED_NAMED(__POUNAME());
        state_1 := 10;
END_CASE
END_METHOD

METHOD PRIVATE Test_StoppedGivesNoOutput
TcUnit.TEST(__POUNAME());
// act
group_3(Run := FALSE);
fb_3(TonIn1 := TRUE);
// assert
AssertEquals_BOOL(Expected := FALSE, Actual := fb_3.TonOut, Message := 'no output while the group is stopped');
AssertEquals_BOOL(Expected := FALSE, Actual := fb_3.IsRunning, Message := 'not running while the group is stopped');
TEST_FINISHED_NAMED(__POUNAME());
END_METHOD

END_FUNCTION_BLOCK

// Tests/User_FB_Tests/T_SafePulse_UserFB_Tests_CFC
    // CFC twin of T_SafePulse_UserFB_Tests: the same tests drawn as CFC diagrams, the way a TwinSAFE project is authored.
    FUNCTION_BLOCK T_SafePulse_UserFB_Tests_CFC EXTENDS T_SafeCfcTestSuite
    VAR
    // Test_PulseForDelayTimeWhileInputHeld
    group_1 : T_SafeGroup;
    fb_1 : T_SafePulse_UserFB(group := group_1) := (Parameters := (DelayTime := T#100MS));
    trigStart_1 : R_TRIG;
    t1_1 : TON;
    t2_1 : TON;
    trig1_1 : R_TRIG;
    trig2_1 : R_TRIG;
    // Test_PulseEndsWhenInputDrops
    group_2 : T_SafeGroup;
    fb_2 : T_SafePulse_UserFB(group := group_2) := (Parameters := (DelayTime := T#100MS));
    // Test_StoppedGivesNoOutput
    group_3 : T_SafeGroup;
    fb_3 : T_SafePulse_UserFB(group := group_3) := (Parameters := (DelayTime := T#100MS));
    // Test_InnerBlocksJoinTheGroup
    group_4 : T_SafeGroup;
    fb_4 : T_SafePulse_UserFB(group := group_4);
END_VAR

Test_PulseForDelayTimeWhileInputHeld();
Test_PulseEndsWhenInputDrops();
Test_StoppedGivesNoOutput();
Test_InnerBlocksJoinTheGroup();

METHOD PRIVATE Test_InnerBlocksJoinTheGroup
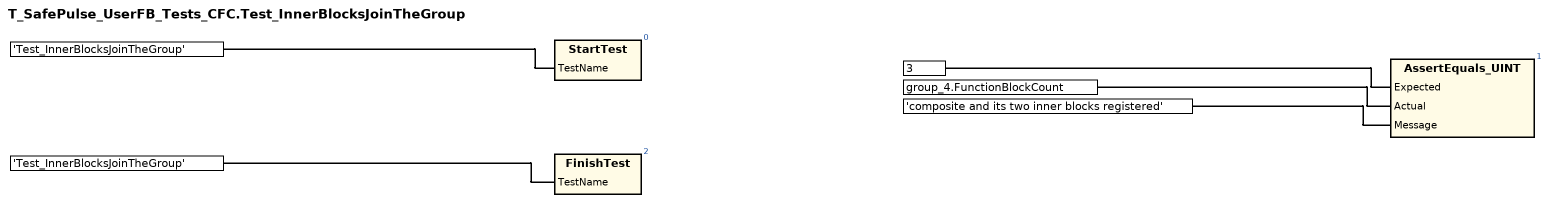
StartTest(TestName := 'Test_InnerBlocksJoinTheGroup');
AssertEquals_UINT(Expected := 3, Actual := group_4.FunctionBlockCount, Message := 'composite and its two inner blocks registered');
FinishTest(TestName := 'Test_InnerBlocksJoinTheGroup');
END_METHOD

METHOD PRIVATE Test_PulseEndsWhenInputDrops
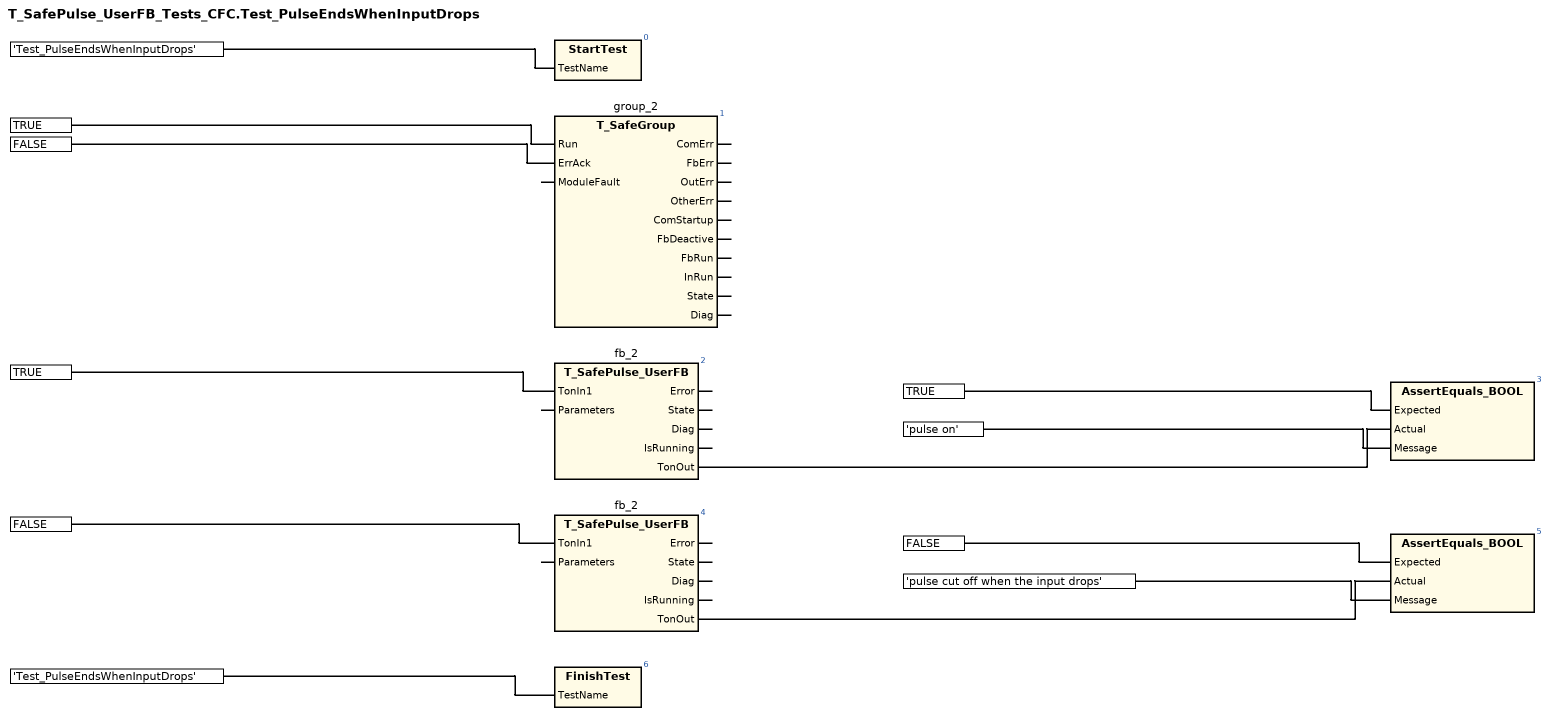
StartTest(TestName := 'Test_PulseEndsWhenInputDrops');
group_2(Run := TRUE, ErrAck := FALSE); // T_SafeGroup
fb_2(TonIn1 := TRUE); // T_SafePulse_UserFB
AssertEquals_BOOL(Expected := TRUE, Actual := fb_2.TonOut, Message := 'pulse on');
fb_2(TonIn1 := FALSE); // T_SafePulse_UserFB
AssertEquals_BOOL(Expected := FALSE, Actual := fb_2.TonOut, Message := 'pulse cut off when the input drops');
FinishTest(TestName := 'Test_PulseEndsWhenInputDrops');
END_METHOD

METHOD PRIVATE Test_PulseForDelayTimeWhileInputHeld
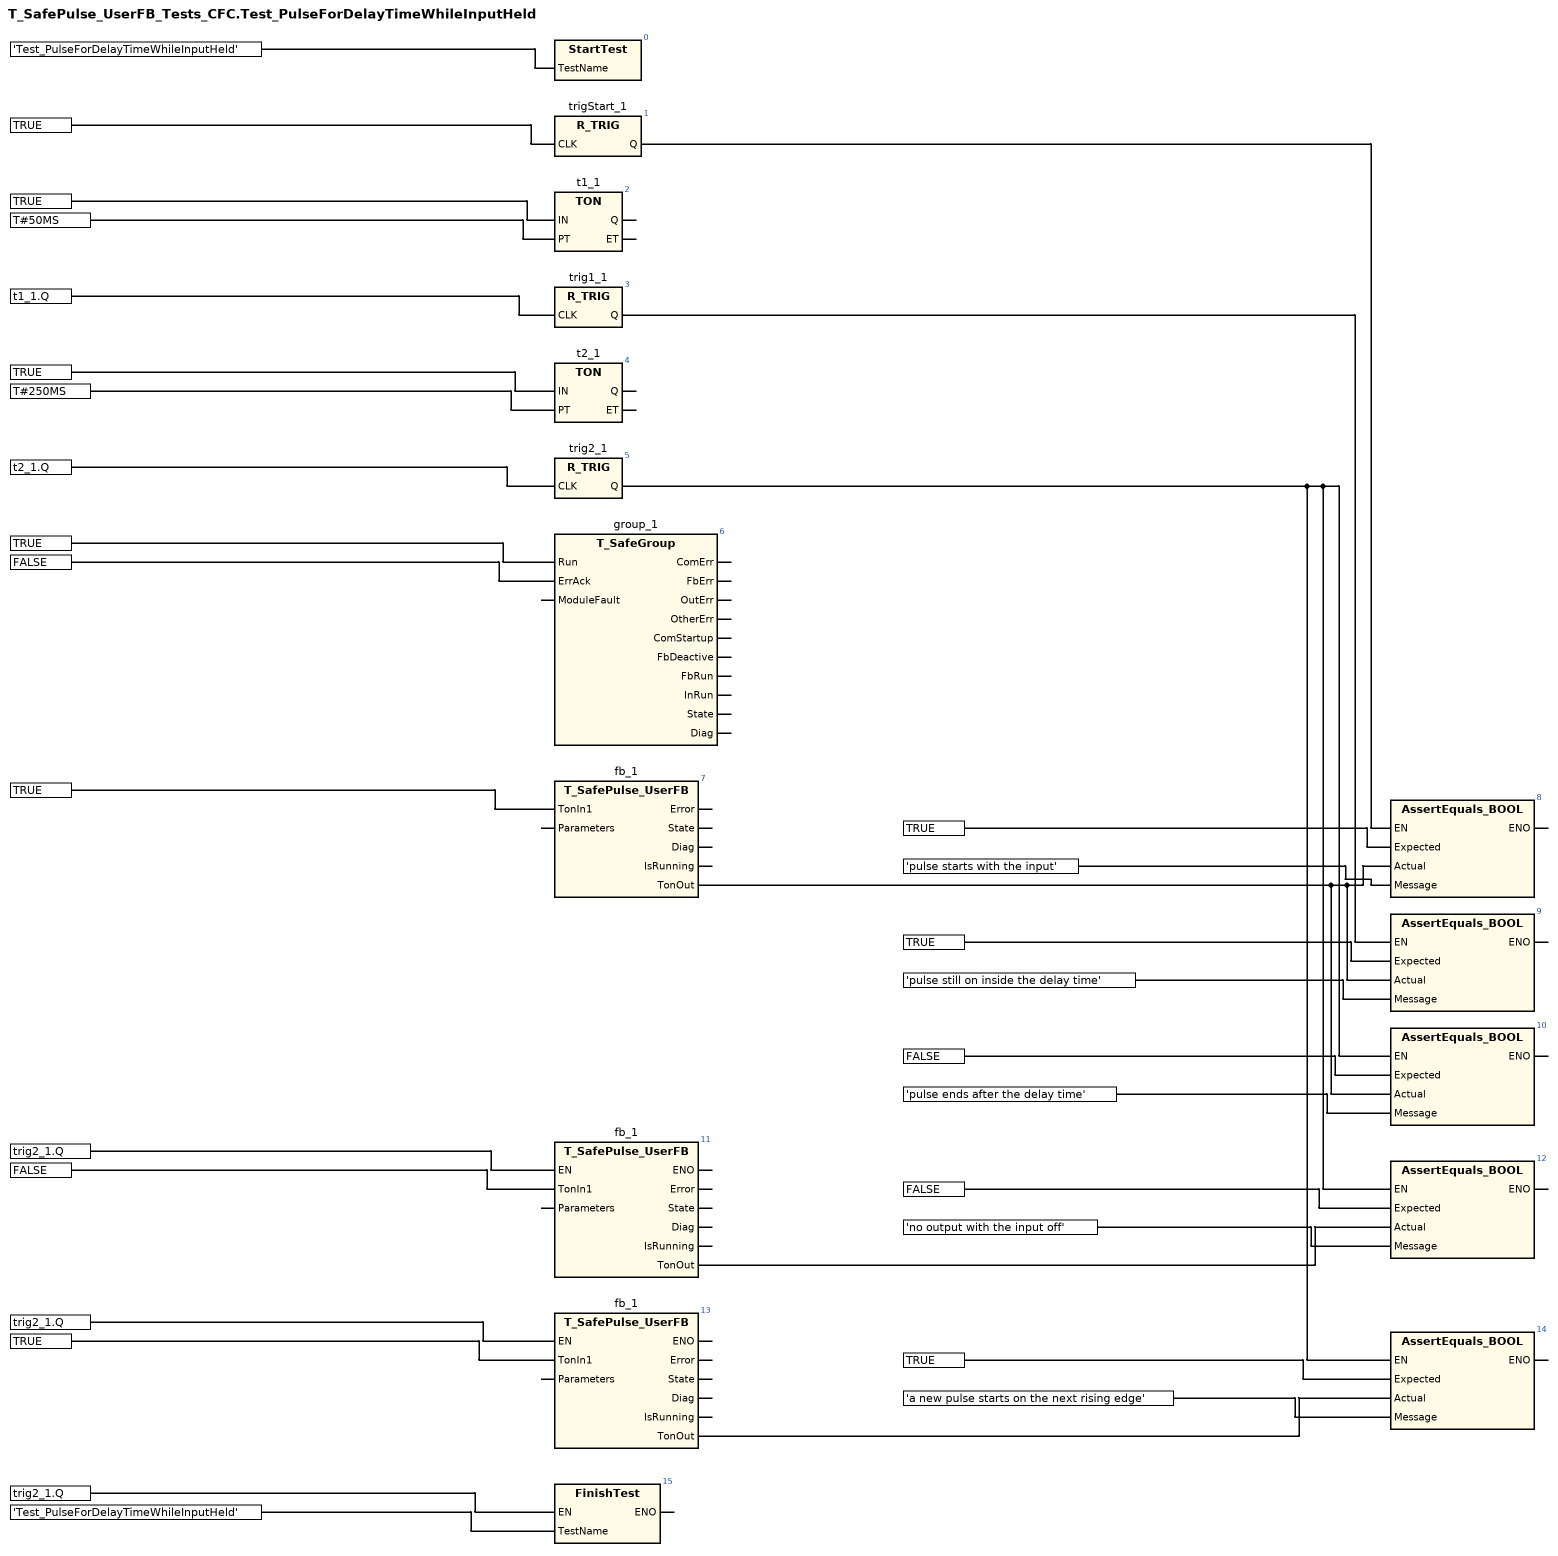
StartTest(TestName := 'Test_PulseForDelayTimeWhileInputHeld');
trigStart_1(CLK := TRUE); // R_TRIG
t1_1(IN := TRUE, PT := T#50MS); // TON
trig1_1(CLK := t1_1.Q); // R_TRIG
t2_1(IN := TRUE, PT := T#250MS); // TON
trig2_1(CLK := t2_1.Q); // R_TRIG
group_1(Run := TRUE, ErrAck := FALSE); // T_SafeGroup
fb_1(TonIn1 := TRUE); // T_SafePulse_UserFB
IF trigStart_1.Q THEN AssertEquals_BOOL(Expected := TRUE, Actual := fb_1.TonOut, Message := 'pulse starts with the input'); END_IF
IF trig1_1.Q THEN AssertEquals_BOOL(Expected := TRUE, Actual := fb_1.TonOut, Message := 'pulse still on inside the delay time'); END_IF
IF trig2_1.Q THEN AssertEquals_BOOL(Expected := FALSE, Actual := fb_1.TonOut, Message := 'pulse ends after the delay time'); END_IF
IF trig2_1.Q THEN
    fb_1(TonIn1 := FALSE); // T_SafePulse_UserFB
END_IF
IF trig2_1.Q THEN AssertEquals_BOOL(Expected := FALSE, Actual := fb_1.TonOut, Message := 'no output with the input off'); END_IF
IF trig2_1.Q THEN
    fb_1(TonIn1 := TRUE); // T_SafePulse_UserFB
END_IF
IF trig2_1.Q THEN AssertEquals_BOOL(Expected := TRUE, Actual := fb_1.TonOut, Message := 'a new pulse starts on the next rising edge'); END_IF
IF trig2_1.Q THEN FinishTest(TestName := 'Test_PulseForDelayTimeWhileInputHeld'); END_IF
END_METHOD

METHOD PRIVATE Test_StoppedGivesNoOutput
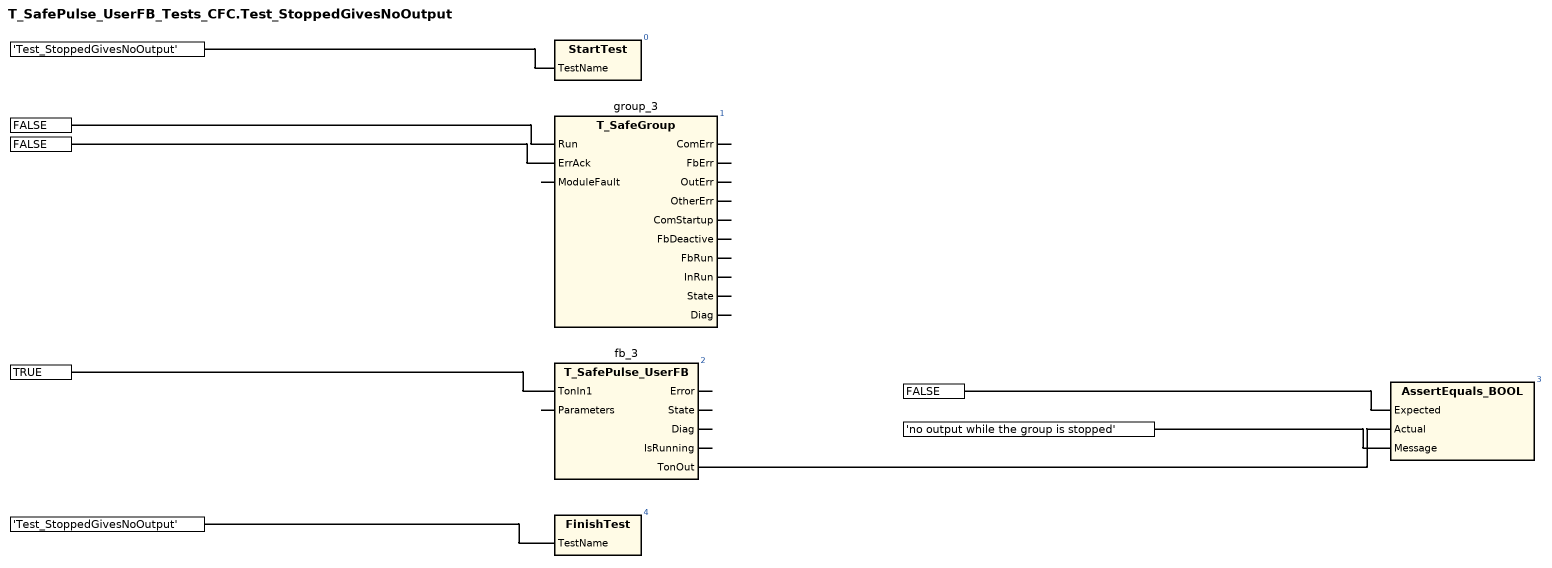
StartTest(TestName := 'Test_StoppedGivesNoOutput');
group_3(Run := FALSE, ErrAck := FALSE); // T_SafeGroup
fb_3(TonIn1 := TRUE); // T_SafePulse_UserFB
AssertEquals_BOOL(Expected := FALSE, Actual := fb_3.TonOut, Message := 'no output while the group is stopped');
FinishTest(TestName := 'Test_StoppedGivesNoOutput');
END_METHOD

END_FUNCTION_BLOCK

// Tests/T_SafeCfcTestSuite
// Base of the CFC test suites. TcUnit's TEST and TEST_FINISHED_NAMED are functions without a return
// type, which a CFC box cannot call (the editor insists on a return pin), so the diagrams call these
// two methods instead. Everything else comes from TcUnit.FB_TestSuite.
FUNCTION_BLOCK ABSTRACT T_SafeCfcTestSuite EXTENDS TcUnit.FB_TestSuite

// Marks a test as finished (TcUnit.TEST_FINISHED_NAMED).
METHOD PROTECTED FinishTest
VAR_INPUT
    TestName : T_MaxString;
END_VAR
TcUnit.TEST_FINISHED_NAMED(TestName);
END_METHOD

// Marks the start of a test (TcUnit.TEST). Call it first in every test method, every cycle.
METHOD PROTECTED StartTest
VAR_INPUT
    TestName : T_MaxString;
END_VAR
TcUnit.TEST(TestName);
END_METHOD

END_FUNCTION_BLOCK

// Tests/User_FB_Tests/T_SafeRTrig_UserFB_Tests
// Tests of the example user FB T_SafeRTrig_UserFB: Trigger is on for one cycle on the rising edge of Signal.
FUNCTION_BLOCK T_SafeRTrig_UserFB_Tests EXTENDS TcUnit.FB_TestSuite
VAR
    // Test_TriggerForOneCycleOnRisingEdge
    group_1 : T_SafeGroup;
    fb_1 : T_SafeRTrig_UserFB(group := group_1);
    // Test_StoppedGivesNoOutput
    group_2 : T_SafeGroup;
    fb_2 : T_SafeRTrig_UserFB(group := group_2);
    // Test_InnerBlocksJoinTheGroup
    group_3 : T_SafeGroup;
    fb_3 : T_SafeRTrig_UserFB(group := group_3);
END_VAR

Test_TriggerForOneCycleOnRisingEdge();
Test_StoppedGivesNoOutput();
Test_InnerBlocksJoinTheGroup();

METHOD PRIVATE Test_InnerBlocksJoinTheGroup
TcUnit.TEST(__POUNAME());
// assert: the composite registered itself and passed the group on to its RS and AND
AssertEquals_UINT(Expected := 3, Actual := group_3.FunctionBlockCount, Message := 'composite and its two inner blocks registered');
TEST_FINISHED_NAMED(__POUNAME());
END_METHOD

METHOD PRIVATE Test_StoppedGivesNoOutput
TcUnit.TEST(__POUNAME());
// act
group_2(Run := FALSE);
fb_2(Signal := TRUE);
// assert
AssertEquals_BOOL(Expected := FALSE, Actual := fb_2.Trigger, Message := 'no output while the group is stopped');
AssertEquals_BOOL(Expected := FALSE, Actual := fb_2.IsRunning, Message := 'not running while the group is stopped');
TEST_FINISHED_NAMED(__POUNAME());
END_METHOD

METHOD PRIVATE Test_TriggerForOneCycleOnRisingEdge
TcUnit.TEST(__POUNAME());
// act / assert
group_1(Run := TRUE);
fb_1(Signal := FALSE);
AssertEquals_BOOL(Expected := FALSE, Actual := fb_1.Trigger, Message := 'no trigger while the signal is off');
AssertEquals_BOOL(Expected := TRUE, Actual := fb_1.IsRunning, Message := 'reports Run to the group while it runs');
fb_1(Signal := TRUE);
AssertEquals_BOOL(Expected := TRUE, Actual := fb_1.Trigger, Message := 'trigger on the rising edge');
fb_1(Signal := TRUE);
AssertEquals_BOOL(Expected := FALSE, Actual := fb_1.Trigger, Message := 'trigger lasts one cycle');
fb_1(Signal := FALSE);
AssertEquals_BOOL(Expected := FALSE, Actual := fb_1.Trigger, Message := 'no trigger on the falling edge');
fb_1(Signal := TRUE);
AssertEquals_BOOL(Expected := TRUE, Actual := fb_1.Trigger, Message := 'triggers again on the next rising edge');
TEST_FINISHED_NAMED(__POUNAME());
END_METHOD

END_FUNCTION_BLOCK

// Tests/User_FB_Tests/T_SafeRTrig_UserFB_Tests_CFC
    // CFC twin of T_SafeRTrig_UserFB_Tests: the same tests drawn as CFC diagrams, the way a TwinSAFE project is authored.
    FUNCTION_BLOCK T_SafeRTrig_UserFB_Tests_CFC EXTENDS T_SafeCfcTestSuite
    VAR
    // Test_TriggerForOneCycleOnRisingEdge
    group_1 : T_SafeGroup;
    fb_1 : T_SafeRTrig_UserFB(group := group_1);
    // Test_StoppedGivesNoOutput
    group_2 : T_SafeGroup;
    fb_2 : T_SafeRTrig_UserFB(group := group_2);
    // Test_InnerBlocksJoinTheGroup
    group_3 : T_SafeGroup;
    fb_3 : T_SafeRTrig_UserFB(group := group_3);
END_VAR

Test_TriggerForOneCycleOnRisingEdge();
Test_StoppedGivesNoOutput();
Test_InnerBlocksJoinTheGroup();

METHOD PRIVATE Test_InnerBlocksJoinTheGroup
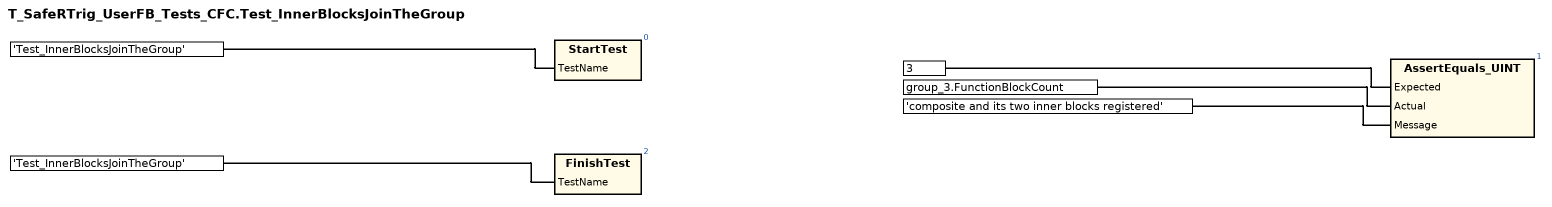
StartTest(TestName := 'Test_InnerBlocksJoinTheGroup');
AssertEquals_UINT(Expected := 3, Actual := group_3.FunctionBlockCount, Message := 'composite and its two inner blocks registered');
FinishTest(TestName := 'Test_InnerBlocksJoinTheGroup');
END_METHOD

METHOD PRIVATE Test_StoppedGivesNoOutput
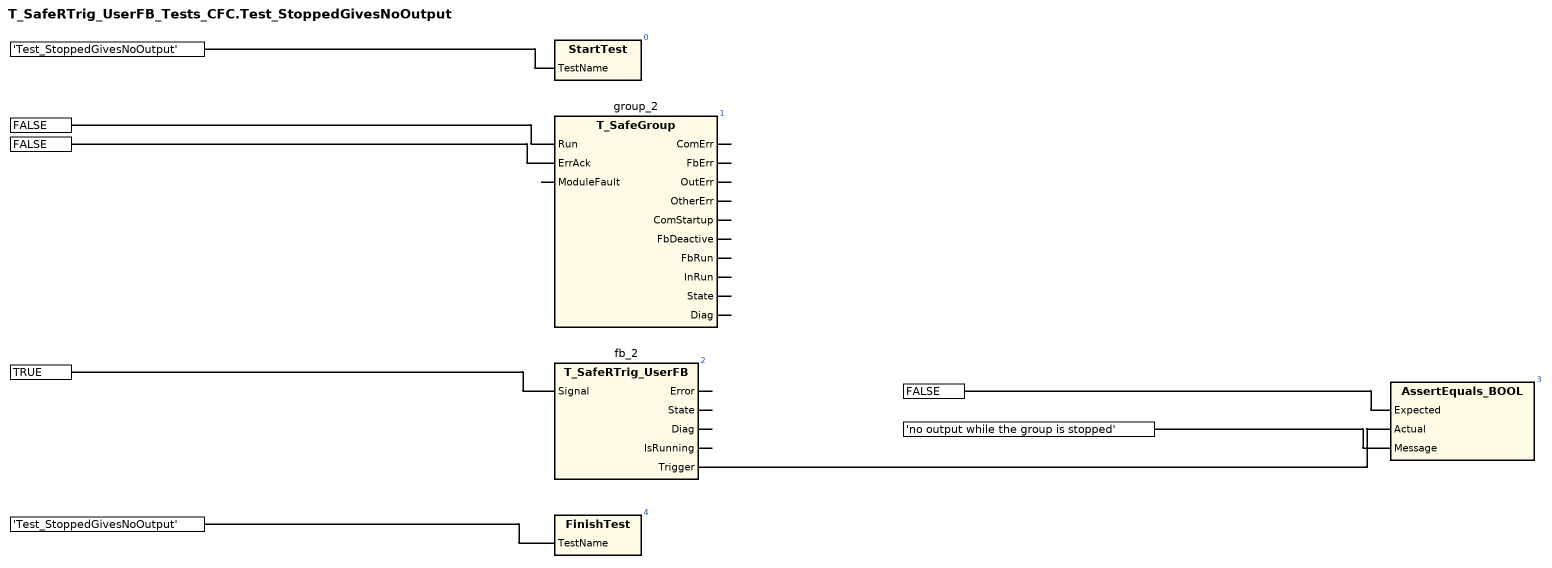
StartTest(TestName := 'Test_StoppedGivesNoOutput');
group_2(Run := FALSE, ErrAck := FALSE); // T_SafeGroup
fb_2(Signal := TRUE); // T_SafeRTrig_UserFB
AssertEquals_BOOL(Expected := FALSE, Actual := fb_2.Trigger, Message := 'no output while the group is stopped');
FinishTest(TestName := 'Test_StoppedGivesNoOutput');
END_METHOD

METHOD PRIVATE Test_TriggerForOneCycleOnRisingEdge
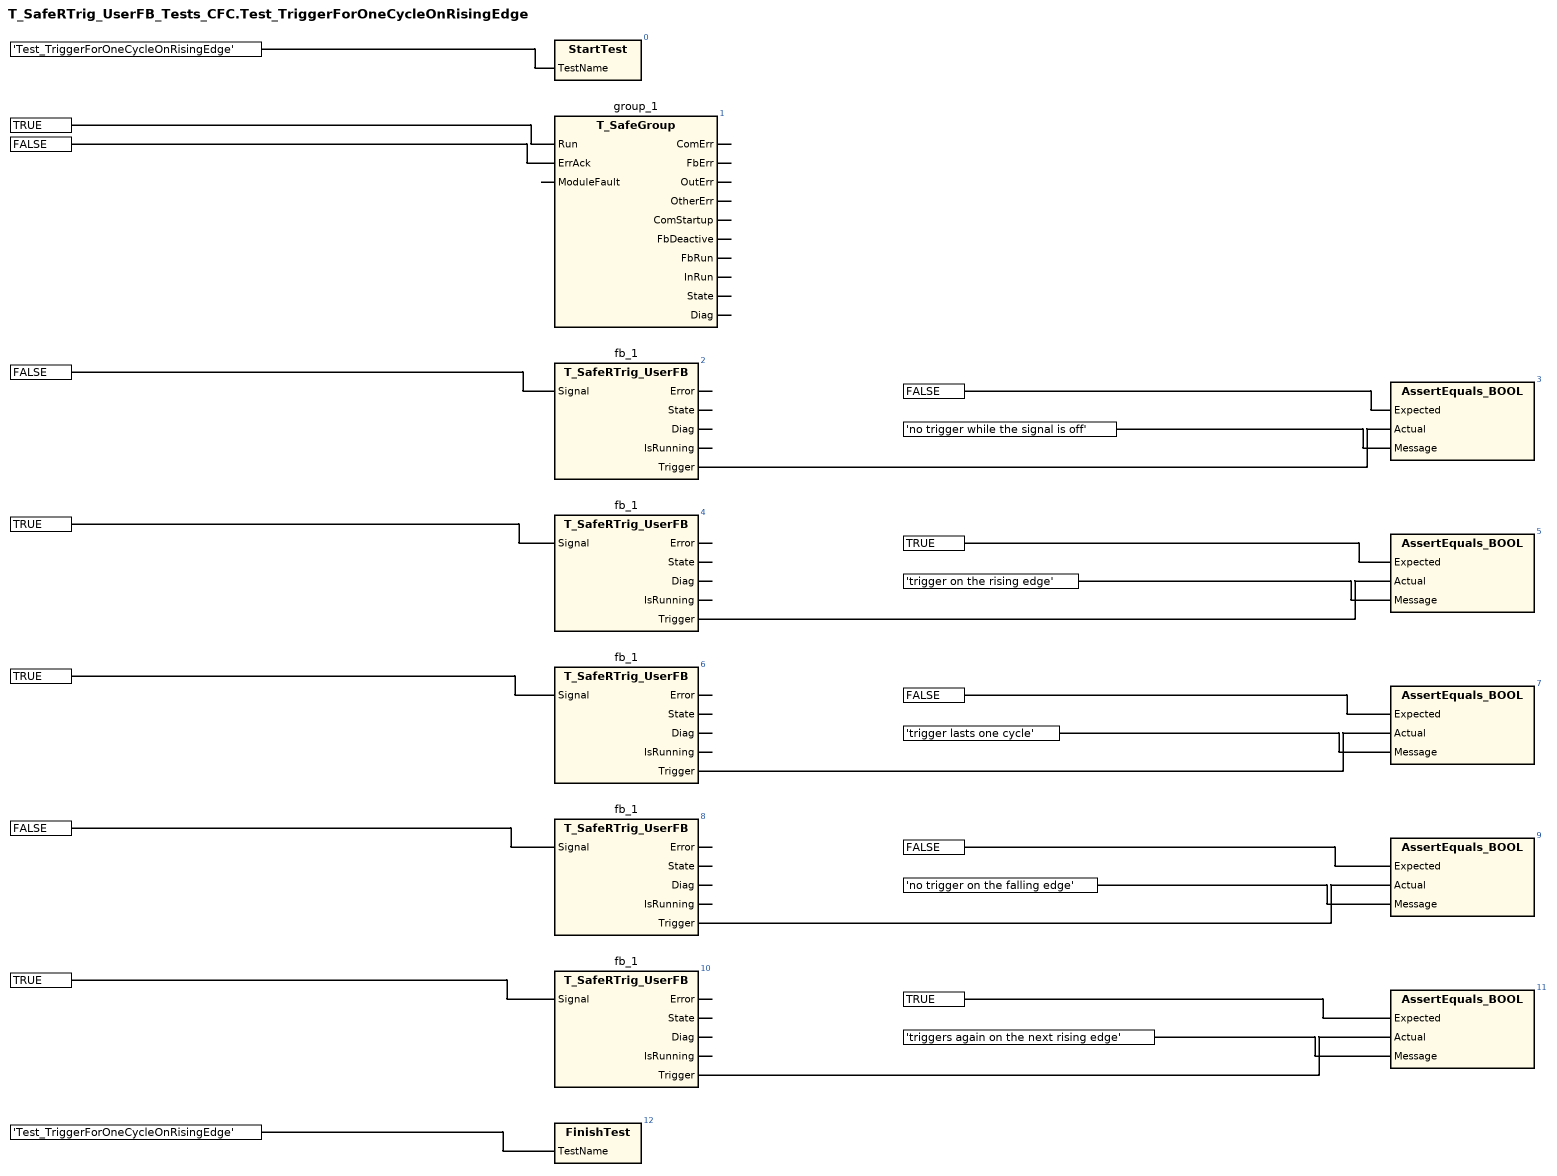
StartTest(TestName := 'Test_TriggerForOneCycleOnRisingEdge');
group_1(Run := TRUE, ErrAck := FALSE); // T_SafeGroup
fb_1(Signal := FALSE); // T_SafeRTrig_UserFB
AssertEquals_BOOL(Expected := FALSE, Actual := fb_1.Trigger, Message := 'no trigger while the signal is off');
fb_1(Signal := TRUE); // T_SafeRTrig_UserFB
AssertEquals_BOOL(Expected := TRUE, Actual := fb_1.Trigger, Message := 'trigger on the rising edge');
fb_1(Signal := TRUE); // T_SafeRTrig_UserFB
AssertEquals_BOOL(Expected := FALSE, Actual := fb_1.Trigger, Message := 'trigger lasts one cycle');
fb_1(Signal := FALSE); // T_SafeRTrig_UserFB
AssertEquals_BOOL(Expected := FALSE, Actual := fb_1.Trigger, Message := 'no trigger on the falling edge');
fb_1(Signal := TRUE); // T_SafeRTrig_UserFB
AssertEquals_BOOL(Expected := TRUE, Actual := fb_1.Trigger, Message := 'triggers again on the next rising edge');
FinishTest(TestName := 'Test_TriggerForOneCycleOnRisingEdge');
END_METHOD

END_FUNCTION_BLOCK

// Tests/PRG_TestRunner
// Runs every TcUnit test suite in the library.
PROGRAM PRG_TestRunner
VAR
    safeAndTests                    : T_SafeAnd_Tests;
    safeInputPairTests              : T_SafeInputPair_Tests;
    safeOrTests                     : T_SafeOr_Tests;
    safeXorTests                    : T_SafeXor_Tests;
    safeDecoupleTests               : T_SafeDecouple_Tests;
    safeOpModeTests                 : T_SafeOpMode_Tests;
    safeRsTests                     : T_SafeRs_Tests;
    safeSrTests                     : T_SafeSr_Tests;
    safeTonTests                    : T_SafeTon_Tests;
    safeTofTests                    : T_SafeTof_Tests;
    safeEdmTests                    : T_SafeEdm_Tests;
    safeEStopTests                  : T_SafeEStop_Tests;
    safeMonTests                    : T_SafeMon_Tests;
    safeTwoHandTests                : T_SafeTwoHand_Tests;
    safeMutingTests                 : T_SafeMuting_Tests;
    safeConnectionTests             : T_SafeConnection_Tests;
    safeInputTerminal8Tests         : T_SafeInputTerminal8_Tests;
    safeOutputTerminal2Tests        : T_SafeOutputTerminal2_Tests;
    safeConnShutdownTests           : T_SafeConnShutdown_Tests;
    safeGroupTests                  : T_SafeGroup_Tests;
    safePulseUserFbTests            : T_SafePulse_UserFB_Tests;
    safeRTrigUserFbTests            : T_SafeRTrig_UserFB_Tests;

    // CFC twins of the suites above
    safeAndTestsCfc                 : T_SafeAnd_Tests_CFC;
    safeInputPairTestsCfc           : T_SafeInputPair_Tests_CFC;
    safeOrTestsCfc                  : T_SafeOr_Tests_CFC;
    safeXorTestsCfc                 : T_SafeXor_Tests_CFC;
    safeDecoupleTestsCfc            : T_SafeDecouple_Tests_CFC;
    safeOpModeTestsCfc              : T_SafeOpMode_Tests_CFC;
    safeRsTestsCfc                  : T_SafeRs_Tests_CFC;
    safeSrTestsCfc                  : T_SafeSr_Tests_CFC;
    safeTonTestsCfc                 : T_SafeTon_Tests_CFC;
    safeTofTestsCfc                 : T_SafeTof_Tests_CFC;
    safeEdmTestsCfc                 : T_SafeEdm_Tests_CFC;
    safeEStopTestsCfc               : T_SafeEStop_Tests_CFC;
    safeMonTestsCfc                 : T_SafeMon_Tests_CFC;
    safeTwoHandTestsCfc             : T_SafeTwoHand_Tests_CFC;
    safeMutingTestsCfc              : T_SafeMuting_Tests_CFC;
    safeConnectionTestsCfc          : T_SafeConnection_Tests_CFC;
    safeConnShutdownTestsCfc        : T_SafeConnShutdown_Tests_CFC;
    safeGroupTestsCfc               : T_SafeGroup_Tests_CFC;
    safePulseUserFbTestsCfc         : T_SafePulse_UserFB_Tests_CFC;
    safeRTrigUserFbTestsCfc         : T_SafeRTrig_UserFB_Tests_CFC;
END_VAR

// Intecre.Utilities logs nothing until a project sets LogConfig.LogLevel; Error lets the
// refused-configuration lines of the configuration tests through to the TwinCAT log.
LogConfig.LogLevel := E_LogSeverity.Error;
TcUnit.RUN();

END_PROGRAM

// Tests/T_SafeAnd_Tests
FUNCTION_BLOCK T_SafeAnd_Tests EXTENDS TcUnit.FB_TestSuite
VAR
    // Test_AllConnectedInputsTrueGivesRun
    group_1 : T_SafeGroup;
    fb_1 : T_SafeAnd(group := group_1);
    // Test_OneInputFalseGivesSafe
    group_2 : T_SafeGroup;
    fb_2 : T_SafeAnd(group := group_2);
    // Test_UnconnectedInputsIgnoredAndMakeContactNegated
    group_3 : T_SafeGroup;
    fb_3 : T_SafeAnd(group := group_3) := (Parameters := (In2MakeContact := TRUE));
    // Test_StoppedGivesNoOutput
    group_4 : T_SafeGroup;
    fb_4 : T_SafeAnd(group := group_4);
    // Test_OneConnectedInputIsRefused
    group_5 : T_SafeGroup;
    fb_5 : T_SafeAnd(group := group_5);
    // Test_RaiseOnRefusedConfigurationStopsHard
    group_6 : T_SafeGroup;
    fb_6 : T_SafeAnd(group := group_6);
END_VAR

Test_AllConnectedInputsTrueGivesRun();
Test_OneInputFalseGivesSafe();
Test_UnconnectedInputsIgnoredAndMakeContactNegated();
Test_StoppedGivesNoOutput();
Test_OneConnectedInputIsRefused();
Test_RaiseOnRefusedConfigurationStopsHard();

METHOD PRIVATE Test_AllConnectedInputsTrueGivesRun
TcUnit.TEST(__POUNAME());
// act
group_1(Run := TRUE);
fb_1(AndIn1 := TRUE, AndIn2 := TRUE);
// assert
AssertEquals_BOOL(Expected := TRUE, Actual := fb_1.AndOut, Message := 'output on when all connected inputs are 1');
AssertEquals_BYTE(Expected := TO_BYTE(E_SafeFbState.Run), Actual := fb_1.State, Message := 'state RUN');
TEST_FINISHED_NAMED(__POUNAME());
END_METHOD

METHOD PRIVATE Test_OneConnectedInputIsRefused
TcUnit.TEST(__POUNAME());
// arrange / act: AndIn1 is the only connected input, which the Safety Editor refuses
group_5(Run := TRUE);
fb_5(AndIn1 := TRUE);
group_5(Run := TRUE);
fb_5(AndIn1 := TRUE);
// assert
AssertEquals_BOOL(Expected := TRUE, Actual := fb_5.Error, Message := 'configuration error reported');
AssertEquals_BYTE(Expected := TO_BYTE(E_SafeFbState.Error), Actual := fb_5.State, Message := 'state ERROR');
AssertEquals_WORD(Expected := WORD#16#8000, Actual := fb_5.Diag, Message := 'diag bit 15 configuration refused');
AssertEquals_BOOL(Expected := FALSE, Actual := fb_5.AndOut, Message := 'AndOut stays at its safe value');
AssertEquals_BOOL(Expected := TRUE, Actual := group_5.FbErr, Message := 'the group sees an FB error');
// act: ErrAck 0 -> 1 -> 0 does not clear a configuration error
group_5(Run := TRUE, ErrAck := TRUE);
fb_5(AndIn1 := TRUE);
group_5(Run := TRUE, ErrAck := TRUE);
fb_5(AndIn1 := TRUE);
group_5(Run := TRUE, ErrAck := FALSE);
fb_5(AndIn1 := TRUE);
AssertEquals_BOOL(Expected := TRUE, Actual := fb_5.Error, Message := 'error not acknowledged');
AssertEquals_WORD(Expected := WORD#16#8000, Actual := fb_5.Diag, Message := 'diag bit 15 kept');
TEST_FINISHED_NAMED(__POUNAME());
END_METHOD

METHOD PRIVATE Test_OneInputFalseGivesSafe
TcUnit.TEST(__POUNAME());
// act
group_2(Run := TRUE);
fb_2(AndIn1 := TRUE, AndIn2 := FALSE);
// assert
AssertEquals_BOOL(Expected := FALSE, Actual := fb_2.AndOut, Message := 'output off when a connected input is 0');
AssertEquals_BYTE(Expected := TO_BYTE(E_SafeFbState.Safe), Actual := fb_2.State, Message := 'state SAFE');
TEST_FINISHED_NAMED(__POUNAME());
END_METHOD

METHOD PRIVATE Test_RaiseOnRefusedConfigurationStopsHard
VAR
    exc : __SYSTEM.ExceptionCode;
    caught : __SYSTEM.ExceptionCode;
END_VAR
TcUnit.TEST(__POUNAME());
// arrange: a one-input AND, the group's opt-in hard stop switched on for this call only
caught := __SYSTEM.ExceptionCode.RTSEXCPT_NOEXCEPTION;
group_6.RaiseOnRefusedConfiguration := TRUE;
// act
__TRY
    group_6(Run := TRUE);
    fb_6(AndIn1 := TRUE);
__CATCH(exc)
    caught := exc;
__FINALLY
    group_6.RaiseOnRefusedConfiguration := FALSE;
__ENDTRY
// assert: the code given to F_RaiseException does not reach __CATCH on TwinCAT 3.1 4026 (the x64
// usermode runtime delivered 16#E8940001 instead of RTSEXCPT_IO_CONFIG_ERROR), so only the arrival
// of an exception is checked; the block's own outputs carry the reason
AssertEquals_BOOL(Expected := TRUE, Actual := (caught <> __SYSTEM.ExceptionCode.RTSEXCPT_NOEXCEPTION), Message := 'an exception was raised and caught');
AssertEquals_BOOL(Expected := TRUE, Actual := fb_6.Error, Message := 'error reported before the exception');
AssertEquals_BYTE(Expected := TO_BYTE(E_SafeFbState.Error), Actual := fb_6.State, Message := 'state ERROR');
AssertEquals_WORD(Expected := WORD#16#8000, Actual := fb_6.Diag, Message := 'diag bit 15 configuration refused');
TEST_FINISHED_NAMED(__POUNAME());
END_METHOD

METHOD PRIVATE Test_StoppedGivesNoOutput
TcUnit.TEST(__POUNAME());
// act
group_4(Run := FALSE);
fb_4(AndIn1 := TRUE, AndIn2 := TRUE);
// assert
AssertEquals_BOOL(Expected := FALSE, Actual := fb_4.AndOut, Message := 'no output while the group is stopped');
AssertEquals_BYTE(Expected := TO_BYTE(E_SafeFbState.Stop), Actual := fb_4.State, Message := 'state STOP');
TEST_FINISHED_NAMED(__POUNAME());
END_METHOD

METHOD PRIVATE Test_UnconnectedInputsIgnoredAndMakeContactNegated
TcUnit.TEST(__POUNAME());
// act: AndIn3..8 unconnected, AndIn2 make contact at 0 (released)
group_3(Run := TRUE);
fb_3(AndIn1 := TRUE, AndIn2 := FALSE);
// assert
AssertEquals_BOOL(Expected := TRUE, Actual := fb_3.AndOut, Message := 'unconnected inputs ignored, make contact negated');
TEST_FINISHED_NAMED(__POUNAME());
END_METHOD

END_FUNCTION_BLOCK

// Tests/T_SafeInputPair_Tests
FUNCTION_BLOCK T_SafeInputPair_Tests EXTENDS TcUnit.FB_TestSuite
VAR
    // Test_DiscrepancyErrorAfterTimeoutAndResetAfterSafeInputs
    pair_5 : T_SafeInputPair;
    state_5 : INT := 10;
    waitTimer_5 : TON;
END_VAR

Test_InactivePairNeverRequestsSafeState();
Test_BreakContactRequestsSafeStateOnZero();
Test_MakeContactRequestsSafeStateOnOne();
Test_TwoChannelRequestsSafeStateIfEitherChannelLow();
Test_DiscrepancyErrorAfterTimeoutAndResetAfterSafeInputs();

METHOD PRIVATE Test_BreakContactRequestsSafeStateOnZero
VAR
    pair : T_SafeInputPair;
END_VAR
TcUnit.TEST(__POUNAME());
// act
pair(In1 := FALSE, Active1 := TRUE, Monitor := TRUE);
// assert
AssertEquals_BOOL(Expected := TRUE, Actual := pair.SafeStateRequested, Message := 'break contact at 0 must request the safe state');
pair(In1 := TRUE, Active1 := TRUE, Monitor := TRUE);
AssertEquals_BOOL(Expected := FALSE, Actual := pair.SafeStateRequested, Message := 'break contact at 1 must not request the safe state');
TEST_FINISHED_NAMED(__POUNAME());
END_METHOD

METHOD PRIVATE Test_DiscrepancyErrorAfterTimeoutAndResetAfterSafeInputs
TcUnit.TEST(__POUNAME());
waitTimer_5();

CASE state_5 OF
    10:
        // arrange
        state_5 := 20;
        waitTimer_5(IN := TRUE, PT := T#50MS);
    20:
        // act: channels disagree for less than the discrepancy time
        pair_5(
            In1 := TRUE,
            In2 := FALSE,
            Active1 := TRUE,
            Active2 := TRUE,
            Monitor := TRUE,
            SafeInputsAfterDiscError := TRUE,
            DiscrepancyTime := T#100MS
        );

        IF NOT waitTimer_5.Q THEN
            RETURN;
        END_IF

        waitTimer_5(IN := FALSE);
        // assert
        AssertEquals_BOOL(Expected := FALSE, Actual := pair_5.DiscrepancyError, Message := 'no error before the discrepancy time');
        state_5 := 30;
        waitTimer_5(IN := TRUE, PT := T#200MS);
    30:
        pair_5(
            In1 := TRUE,
            In2 := FALSE,
            Active1 := TRUE,
            Active2 := TRUE,
            Monitor := TRUE,
            SafeInputsAfterDiscError := TRUE,
            DiscrepancyTime := T#100MS
        );

        IF NOT waitTimer_5.Q THEN
            RETURN;
        END_IF

        waitTimer_5(IN := FALSE);
        // assert
        AssertEquals_BOOL(Expected := TRUE, Actual := pair_5.DiscrepancyError, Message := 'error after the discrepancy time');
        AssertEquals_BOOL(Expected := TRUE, Actual := pair_5.AwaitingSafeInputs, Message := 'error waits for both channels safe');
        // act: acknowledge while a channel is still high
        pair_5(
            In1 := TRUE,
            In2 := FALSE,
            Active1 := TRUE,
            Active2 := TRUE,
            Monitor := TRUE,
            SafeInputsAfterDiscError := TRUE,
            DiscrepancyTime := T#100MS,
            Acknowledge := TRUE
        );

        AssertEquals_BOOL(Expected := TRUE, Actual := pair_5.DiscrepancyError, Message := 'acknowledge refused while a channel is still high');
        // act: both channels safe, then acknowledge
        pair_5(
            In1 := FALSE,
            In2 := FALSE,
            Active1 := TRUE,
            Active2 := TRUE,
            Monitor := TRUE,
            SafeInputsAfterDiscError := TRUE,
            DiscrepancyTime := T#100MS,
            Acknowledge := TRUE
        );

        AssertEquals_BOOL(Expected := FALSE, Actual := pair_5.DiscrepancyError, Message := 'error cleared once both channels were safe');
        TEST_FINISHED_NAMED(__POUNAME());
        state_5 := 10;
END_CASE
END_METHOD

METHOD PRIVATE Test_InactivePairNeverRequestsSafeState
VAR
    pair : T_SafeInputPair;
END_VAR
TcUnit.TEST(__POUNAME());
// act
pair(In1 := FALSE, In2 := FALSE, Active1 := FALSE, Active2 := FALSE, Monitor := TRUE);
// assert
AssertEquals_BOOL(Expected := FALSE, Actual := pair.SafeStateRequested, Message := 'inactive pair must not request the safe state');
AssertEquals_BOOL(Expected := FALSE, Actual := pair.IsActive, Message := 'pair should be inactive');
TEST_FINISHED_NAMED(__POUNAME());
END_METHOD

METHOD PRIVATE Test_MakeContactRequestsSafeStateOnOne
VAR
    pair : T_SafeInputPair;
END_VAR
TcUnit.TEST(__POUNAME());
// act
pair(In1 := TRUE, Active1 := TRUE, MakeContact1 := TRUE, Monitor := TRUE);
// assert
AssertEquals_BOOL(Expected := TRUE, Actual := pair.SafeStateRequested, Message := 'make contact at 1 must request the safe state');
TEST_FINISHED_NAMED(__POUNAME());
END_METHOD

METHOD PRIVATE Test_TwoChannelRequestsSafeStateIfEitherChannelLow
VAR
    pair : T_SafeInputPair;
END_VAR
TcUnit.TEST(__POUNAME());
// act
pair(
    In1 := TRUE,
    In2 := FALSE,
    Active1 := TRUE,
    Active2 := TRUE,
    Monitor := TRUE,
    SafeInputsAfterDiscError := TRUE
);

// assert
AssertEquals_BOOL(Expected := TRUE, Actual := pair.SafeStateRequested, Message := 'one low channel must request the safe state');
AssertEquals_BOOL(Expected := FALSE, Actual := pair.DiscrepancyError, Message := 'no discrepancy monitoring without a discrepancy time');
pair(
    In1 := TRUE,
    In2 := TRUE,
    Active1 := TRUE,
    Active2 := TRUE,
    Monitor := TRUE,
    SafeInputsAfterDiscError := TRUE
);

AssertEquals_BOOL(Expected := FALSE, Actual := pair.SafeStateRequested, Message := 'both channels high must not request the safe state');
TEST_FINISHED_NAMED(__POUNAME());
END_METHOD

END_FUNCTION_BLOCK

// Tests/T_SafeOr_Tests
FUNCTION_BLOCK T_SafeOr_Tests EXTENDS TcUnit.FB_TestSuite
VAR
    // Test_AnyConnectedInputTrueGivesRun
    group_1 : T_SafeGroup;
    fb_1 : T_SafeOr(group := group_1);
    // Test_AllFalseGivesSafe
    group_2 : T_SafeGroup;
    fb_2 : T_SafeOr(group := group_2);
    // Test_OneConnectedInputIsRefused
    group_3 : T_SafeGroup;
    fb_3 : T_SafeOr(group := group_3);
END_VAR

Test_AnyConnectedInputTrueGivesRun();
Test_AllFalseGivesSafe();
Test_OneConnectedInputIsRefused();

METHOD PRIVATE Test_AllFalseGivesSafe
TcUnit.TEST(__POUNAME());
// act
group_2(Run := TRUE);
fb_2(OrIn1 := FALSE, OrIn2 := FALSE);
// assert
AssertEquals_BOOL(Expected := FALSE, Actual := fb_2.OrOut, Message := 'output off when all connected inputs are 0');
AssertEquals_BYTE(Expected := TO_BYTE(E_SafeFbState.Safe), Actual := fb_2.State, Message := 'state SAFE');
TEST_FINISHED_NAMED(__POUNAME());
END_METHOD

METHOD PRIVATE Test_AnyConnectedInputTrueGivesRun
TcUnit.TEST(__POUNAME());
// act
group_1(Run := TRUE);
fb_1(OrIn1 := FALSE, OrIn2 := TRUE);
// assert
AssertEquals_BOOL(Expected := TRUE, Actual := fb_1.OrOut, Message := 'output on when any connected input is 1');
TEST_FINISHED_NAMED(__POUNAME());
END_METHOD

METHOD PRIVATE Test_OneConnectedInputIsRefused
TcUnit.TEST(__POUNAME());
// arrange / act: OrIn1 is the only connected input, which the Safety Editor refuses
group_3(Run := TRUE);
fb_3(OrIn1 := TRUE);
group_3(Run := TRUE);
fb_3(OrIn1 := TRUE);
// assert
AssertEquals_BOOL(Expected := TRUE, Actual := fb_3.Error, Message := 'configuration error reported');
AssertEquals_BYTE(Expected := TO_BYTE(E_SafeFbState.Error), Actual := fb_3.State, Message := 'state ERROR');
AssertEquals_WORD(Expected := WORD#16#8000, Actual := fb_3.Diag, Message := 'diag bit 15 configuration refused');
AssertEquals_BOOL(Expected := FALSE, Actual := fb_3.OrOut, Message := 'OrOut stays at its safe value');
AssertEquals_BOOL(Expected := TRUE, Actual := group_3.FbErr, Message := 'the group sees an FB error');
// act: ErrAck 0 -> 1 -> 0 does not clear a configuration error
group_3(Run := TRUE, ErrAck := TRUE);
fb_3(OrIn1 := TRUE);
group_3(Run := TRUE, ErrAck := TRUE);
fb_3(OrIn1 := TRUE);
group_3(Run := TRUE, ErrAck := FALSE);
fb_3(OrIn1 := TRUE);
AssertEquals_BOOL(Expected := TRUE, Actual := fb_3.Error, Message := 'error not acknowledged');
AssertEquals_WORD(Expected := WORD#16#8000, Actual := fb_3.Diag, Message := 'diag bit 15 kept');
TEST_FINISHED_NAMED(__POUNAME());
END_METHOD

END_FUNCTION_BLOCK

// Tests/T_SafeXor_Tests
FUNCTION_BLOCK T_SafeXor_Tests EXTENDS TcUnit.FB_TestSuite
VAR
    // Test_ConnectedPairsAreExclusiveOr
    group_1 : T_SafeGroup;
    fb_1 : T_SafeXor(group := group_1);
END_VAR

Test_ConnectedPairsAreExclusiveOr();

METHOD PRIVATE Test_ConnectedPairsAreExclusiveOr
TcUnit.TEST(__POUNAME());
// act
group_1(Run := TRUE);
fb_1(Xor1In1 := TRUE, Xor2In1 := FALSE);
// assert
AssertEquals_BOOL(Expected := TRUE, Actual := fb_1.XorOut1, Message := 'connected pair 1 XOR');
AssertEquals_BOOL(Expected := FALSE, Actual := fb_1.XorOut2, Message := 'unconnected pair stays 0');
fb_1(Xor1In1 := TRUE, Xor2In1 := TRUE);
AssertEquals_BOOL(Expected := FALSE, Actual := fb_1.XorOut1, Message := 'both inputs 1 gives 0');
TEST_FINISHED_NAMED(__POUNAME());
END_METHOD

END_FUNCTION_BLOCK

// Tests/T_SafeDecouple_Tests
FUNCTION_BLOCK T_SafeDecouple_Tests EXTENDS TcUnit.FB_TestSuite
VAR
    // Test_InputsLoopedToOutputsOnlyWhenRunning
    group_1 : T_SafeGroup;
    fb_1 : T_SafeDecouple(group := group_1);
END_VAR

Test_InputsLoopedToOutputsOnlyWhenRunning();

METHOD PRIVATE Test_InputsLoopedToOutputsOnlyWhenRunning
TcUnit.TEST(__POUNAME());
// act
group_1(Run := TRUE);
fb_1(DecIn3 := TRUE);
// assert
AssertEquals_BOOL(Expected := TRUE, Actual := fb_1.DecOut3, Message := 'input looped to output');
group_1(Run := FALSE);
fb_1(DecIn3 := TRUE);
AssertEquals_BOOL(Expected := FALSE, Actual := fb_1.DecOut3, Message := 'output off while the group is stopped');
TEST_FINISHED_NAMED(__POUNAME());
END_METHOD

END_FUNCTION_BLOCK

// Tests/T_SafeOpMode_Tests
FUNCTION_BLOCK T_SafeOpMode_Tests EXTENDS TcUnit.FB_TestSuite
VAR
    // Test_ExactlyOneInputSelectsOutput
    group_1 : T_SafeGroup;
    fb_1 : T_SafeOpMode(group := group_1);
    // Test_ConnectedRestartRequiresRestartSequence
    group_2 : T_SafeGroup;
    fb_2 : T_SafeOpMode(group := group_2);
    // Test_SlowModeChangeGivesDiscrepancyError
    group_3 : T_SafeGroup;
    fb_3 : T_SafeOpMode(group := group_3) := (Parameters := (DiscrepancyTime := T#100MS));
    state_3 : INT := 10;
    waitTimer_3 : TON;
    // Test_OneConnectedInputIsRefused
    group_4 : T_SafeGroup;
    fb_4 : T_SafeOpMode(group := group_4);
END_VAR

Test_ExactlyOneInputSelectsOutput();
Test_ConnectedRestartRequiresRestartSequence();
Test_SlowModeChangeGivesDiscrepancyError();
Test_OneConnectedInputIsRefused();

METHOD PRIVATE Test_ConnectedRestartRequiresRestartSequence
TcUnit.TEST(__POUNAME());
// act
group_2(Run := TRUE);
fb_2(Restart := FALSE, OpIn1 := TRUE, OpIn2 := FALSE);
group_2(Run := TRUE);
fb_2(Restart := FALSE, OpIn1 := TRUE, OpIn2 := FALSE);
// assert
AssertEquals_BOOL(Expected := FALSE, Actual := fb_2.OpOut1, Message := 'no output before restart');
group_2(Run := TRUE);
fb_2(Restart := TRUE, OpIn1 := TRUE, OpIn2 := FALSE);
AssertEquals_BYTE(Expected := TO_BYTE(E_SafeFbState.Start), Actual := fb_2.State, Message := 'state START while restart held');
group_2(Run := TRUE);
fb_2(Restart := FALSE, OpIn1 := TRUE, OpIn2 := FALSE);
AssertEquals_BOOL(Expected := TRUE, Actual := fb_2.OpOut1, Message := 'output on after restart falling edge');
TEST_FINISHED_NAMED(__POUNAME());
END_METHOD

METHOD PRIVATE Test_ExactlyOneInputSelectsOutput
TcUnit.TEST(__POUNAME());
// act: STOP -> SAFE -> RUN (no Restart connected: automatic)
group_1(Run := TRUE);
fb_1(OpIn1 := FALSE, OpIn2 := TRUE);
group_1(Run := TRUE);
fb_1(OpIn1 := FALSE, OpIn2 := TRUE);
// assert
AssertEquals_BOOL(Expected := TRUE, Actual := fb_1.OpOut2, Message := 'selected mode output on');
AssertEquals_BOOL(Expected := FALSE, Actual := fb_1.OpOut1, Message := 'other outputs off');
AssertEquals_BYTE(Expected := TO_BYTE(E_SafeFbState.Run), Actual := fb_1.State, Message := 'state RUN');
// act: second input also set
group_1(Run := TRUE);
fb_1(OpIn1 := TRUE, OpIn2 := TRUE);
AssertEquals_BOOL(Expected := FALSE, Actual := fb_1.OpOut2, Message := 'all outputs off with two modes selected');
AssertEquals_BYTE(Expected := TO_BYTE(E_SafeFbState.Safe), Actual := fb_1.State, Message := 'state SAFE');
TEST_FINISHED_NAMED(__POUNAME());
END_METHOD

METHOD PRIVATE Test_OneConnectedInputIsRefused
TcUnit.TEST(__POUNAME());
// arrange / act: OpIn1 is the only connected input, which the Safety Editor refuses
group_4(Run := TRUE);
fb_4(OpIn1 := TRUE);
group_4(Run := TRUE);
fb_4(OpIn1 := TRUE);
// assert
AssertEquals_BOOL(Expected := TRUE, Actual := fb_4.Error, Message := 'configuration error reported');
AssertEquals_BYTE(Expected := TO_BYTE(E_SafeFbState.Error), Actual := fb_4.State, Message := 'state ERROR');
AssertEquals_WORD(Expected := WORD#16#8000, Actual := fb_4.Diag, Message := 'diag bit 15 configuration refused');
AssertEquals_BOOL(Expected := FALSE, Actual := fb_4.OpOut1, Message := 'OpOut1 stays at its safe value');
AssertEquals_BOOL(Expected := TRUE, Actual := group_4.FbErr, Message := 'the group sees an FB error');
// act: ErrAck 0 -> 1 -> 0 does not clear a configuration error
group_4(Run := TRUE, ErrAck := TRUE);
fb_4(OpIn1 := TRUE);
group_4(Run := TRUE, ErrAck := TRUE);
fb_4(OpIn1 := TRUE);
group_4(Run := TRUE, ErrAck := FALSE);
fb_4(OpIn1 := TRUE);
AssertEquals_BOOL(Expected := TRUE, Actual := fb_4.Error, Message := 'error not acknowledged');
AssertEquals_WORD(Expected := WORD#16#8000, Actual := fb_4.Diag, Message := 'diag bit 15 kept');
TEST_FINISHED_NAMED(__POUNAME());
END_METHOD

METHOD PRIVATE Test_SlowModeChangeGivesDiscrepancyError
TcUnit.TEST(__POUNAME());
waitTimer_3();

CASE state_3 OF
    10:
        // arrange: mode 1 selected and running
        group_3(Run := TRUE);
        fb_3(OpIn1 := TRUE, OpIn2 := FALSE);
        group_3(Run := TRUE);
        fb_3(OpIn1 := TRUE, OpIn2 := FALSE);
        state_3 := 20;
        waitTimer_3(IN := TRUE, PT := T#250MS);
    20:
        // act: leave mode 1 without selecting another
        group_3(Run := TRUE);
        fb_3(OpIn1 := FALSE, OpIn2 := FALSE);

        IF NOT waitTimer_3.Q THEN
            RETURN;
        END_IF

        waitTimer_3(IN := FALSE);
        // assert
        AssertEquals_BOOL(Expected := TRUE, Actual := fb_3.Error, Message := 'discrepancy error after time without a mode');
        AssertEquals_BYTE(Expected := TO_BYTE(E_SafeFbState.Error), Actual := fb_3.State, Message := 'state ERROR');
        AssertEquals_WORD(Expected := WORD#1, Actual := fb_3.Diag, Message := 'diag bit 0');
        TEST_FINISHED_NAMED(__POUNAME());
        state_3 := 10;
END_CASE
END_METHOD

END_FUNCTION_BLOCK

// Tests/T_SafeRs_Tests
FUNCTION_BLOCK T_SafeRs_Tests EXTENDS TcUnit.FB_TestSuite
VAR
    // Test_ResetDominantLatch
    group_1 : T_SafeGroup;
    fb_1 : T_SafeRs(group := group_1);
    // Test_UnconnectedSetIsRefused
    group_2 : T_SafeGroup;
    fb_2 : T_SafeRs(group := group_2);
END_VAR

Test_ResetDominantLatch();
Test_UnconnectedSetIsRefused();

METHOD PRIVATE Test_ResetDominantLatch
TcUnit.TEST(__POUNAME());
// act / assert
group_1(Run := TRUE);
fb_1(Set := TRUE, Reset := FALSE);
AssertEquals_BOOL(Expected := TRUE, Actual := fb_1.RsOut, Message := 'set');
fb_1(Set := FALSE, Reset := FALSE);
AssertEquals_BOOL(Expected := TRUE, Actual := fb_1.RsOut, Message := 'held');
fb_1(Set := TRUE, Reset := TRUE);
AssertEquals_BOOL(Expected := FALSE, Actual := fb_1.RsOut, Message := 'reset dominant');
TEST_FINISHED_NAMED(__POUNAME());
END_METHOD

METHOD PRIVATE Test_UnconnectedSetIsRefused
TcUnit.TEST(__POUNAME());
// arrange / act: Set is unconnected, which the Safety Editor refuses
group_2(Run := TRUE);
fb_2(Reset := FALSE);
group_2(Run := TRUE);
fb_2(Reset := FALSE);
// assert
AssertEquals_BOOL(Expected := TRUE, Actual := fb_2.Error, Message := 'configuration error reported');
AssertEquals_BYTE(Expected := TO_BYTE(E_SafeFbState.Error), Actual := fb_2.State, Message := 'state ERROR');
AssertEquals_WORD(Expected := WORD#16#8000, Actual := fb_2.Diag, Message := 'diag bit 15 configuration refused');
AssertEquals_BOOL(Expected := FALSE, Actual := fb_2.RsOut, Message := 'RsOut stays at its safe value');
AssertEquals_BOOL(Expected := TRUE, Actual := group_2.FbErr, Message := 'the group sees an FB error');
// act: ErrAck 0 -> 1 -> 0 does not clear a configuration error
group_2(Run := TRUE, ErrAck := TRUE);
fb_2(Reset := FALSE);
group_2(Run := TRUE, ErrAck := TRUE);
fb_2(Reset := FALSE);
group_2(Run := TRUE, ErrAck := FALSE);
fb_2(Reset := FALSE);
AssertEquals_BOOL(Expected := TRUE, Actual := fb_2.Error, Message := 'error not acknowledged');
AssertEquals_WORD(Expected := WORD#16#8000, Actual := fb_2.Diag, Message := 'diag bit 15 kept');
TEST_FINISHED_NAMED(__POUNAME());
END_METHOD

END_FUNCTION_BLOCK

// Tests/T_SafeSr_Tests
FUNCTION_BLOCK T_SafeSr_Tests EXTENDS TcUnit.FB_TestSuite
VAR
    // Test_SetDominantLatch
    group_1 : T_SafeGroup;
    fb_1 : T_SafeSr(group := group_1);
    // Test_UnconnectedResetIsRefused
    group_2 : T_SafeGroup;
    fb_2 : T_SafeSr(group := group_2);
END_VAR

Test_SetDominantLatch();
Test_UnconnectedResetIsRefused();

METHOD PRIVATE Test_SetDominantLatch
TcUnit.TEST(__POUNAME());
// act / assert
group_1(Run := TRUE);
fb_1(Set := TRUE, Reset := TRUE);
AssertEquals_BOOL(Expected := TRUE, Actual := fb_1.SrOut, Message := 'set dominant');
fb_1(Set := FALSE, Reset := TRUE);
AssertEquals_BOOL(Expected := FALSE, Actual := fb_1.SrOut, Message := 'reset');
fb_1(Set := FALSE, Reset := FALSE);
AssertEquals_BOOL(Expected := FALSE, Actual := fb_1.SrOut, Message := 'held');
TEST_FINISHED_NAMED(__POUNAME());
END_METHOD

METHOD PRIVATE Test_UnconnectedResetIsRefused
TcUnit.TEST(__POUNAME());
// arrange / act: Reset is unconnected, which the Safety Editor refuses
group_2(Run := TRUE);
fb_2(Set := TRUE);
group_2(Run := TRUE);
fb_2(Set := TRUE);
// assert
AssertEquals_BOOL(Expected := TRUE, Actual := fb_2.Error, Message := 'configuration error reported');
AssertEquals_BYTE(Expected := TO_BYTE(E_SafeFbState.Error), Actual := fb_2.State, Message := 'state ERROR');
AssertEquals_WORD(Expected := WORD#16#8000, Actual := fb_2.Diag, Message := 'diag bit 15 configuration refused');
AssertEquals_BOOL(Expected := FALSE, Actual := fb_2.SrOut, Message := 'SrOut stays at its safe value');
AssertEquals_BOOL(Expected := TRUE, Actual := group_2.FbErr, Message := 'the group sees an FB error');
// act: ErrAck 0 -> 1 -> 0 does not clear a configuration error
group_2(Run := TRUE, ErrAck := TRUE);
fb_2(Set := TRUE);
group_2(Run := TRUE, ErrAck := TRUE);
fb_2(Set := TRUE);
group_2(Run := TRUE, ErrAck := FALSE);
fb_2(Set := TRUE);
AssertEquals_BOOL(Expected := TRUE, Actual := fb_2.Error, Message := 'error not acknowledged');
AssertEquals_WORD(Expected := WORD#16#8000, Actual := fb_2.Diag, Message := 'diag bit 15 kept');
TEST_FINISHED_NAMED(__POUNAME());
END_METHOD

END_FUNCTION_BLOCK

// Tests/T_SafeTon_Tests
FUNCTION_BLOCK T_SafeTon_Tests EXTENDS TcUnit.FB_TestSuite
VAR
    // Test_OutputDelayedOn
    group_1 : T_SafeGroup;
    fb_1 : T_SafeTon(group := group_1) := (Parameters := (DelayTime := T#100MS));
    state_1 : INT := 10;
    waitTimer_1 : TON;
    // Test_UnconnectedInputIsRefused
    group_2 : T_SafeGroup;
    fb_2 : T_SafeTon(group := group_2);
END_VAR

Test_OutputDelayedOn();
Test_UnconnectedInputIsRefused();

METHOD PRIVATE Test_OutputDelayedOn
TcUnit.TEST(__POUNAME());
waitTimer_1();

CASE state_1 OF
    10:
        // act
        group_1(Run := TRUE);
        fb_1(TonIn1 := TRUE);
        // assert
        AssertEquals_BOOL(Expected := FALSE, Actual := fb_1.TonOut, Message := 'output not yet on');
        AssertEquals_BYTE(Expected := TO_BYTE(E_SafeTonState.DelayIn), Actual := fb_1.State, Message := 'state DELAYIN');
        state_1 := 20;
        waitTimer_1(IN := TRUE, PT := T#200MS);
    20:
        group_1(Run := TRUE);
        fb_1(TonIn1 := TRUE);

        IF NOT waitTimer_1.Q THEN
            RETURN;
        END_IF

        waitTimer_1(IN := FALSE);
        // assert
        AssertEquals_BOOL(Expected := TRUE, Actual := fb_1.TonOut, Message := 'output on after the delay');
        fb_1(TonIn1 := FALSE);
        AssertEquals_BOOL(Expected := FALSE, Actual := fb_1.TonOut, Message := 'output off immediately');
        TEST_FINISHED_NAMED(__POUNAME());
        state_1 := 10;
END_CASE
END_METHOD

METHOD PRIVATE Test_UnconnectedInputIsRefused
TcUnit.TEST(__POUNAME());
// arrange / act: TonIn1 is unconnected, which the Safety Editor refuses
group_2(Run := TRUE);
fb_2();
group_2(Run := TRUE);
fb_2();
// assert
AssertEquals_BOOL(Expected := TRUE, Actual := fb_2.Error, Message := 'configuration error reported');
AssertEquals_BYTE(Expected := TO_BYTE(E_SafeFbState.Error), Actual := fb_2.State, Message := 'state ERROR');
AssertEquals_WORD(Expected := WORD#16#8000, Actual := fb_2.Diag, Message := 'diag bit 15 configuration refused');
AssertEquals_BOOL(Expected := FALSE, Actual := fb_2.TonOut, Message := 'TonOut stays at its safe value');
AssertEquals_BOOL(Expected := TRUE, Actual := group_2.FbErr, Message := 'the group sees an FB error');
// act: ErrAck 0 -> 1 -> 0 does not clear a configuration error
group_2(Run := TRUE, ErrAck := TRUE);
fb_2();
group_2(Run := TRUE, ErrAck := TRUE);
fb_2();
group_2(Run := TRUE, ErrAck := FALSE);
fb_2();
AssertEquals_BOOL(Expected := TRUE, Actual := fb_2.Error, Message := 'error not acknowledged');
AssertEquals_WORD(Expected := WORD#16#8000, Actual := fb_2.Diag, Message := 'diag bit 15 kept');
TEST_FINISHED_NAMED(__POUNAME());
END_METHOD

END_FUNCTION_BLOCK

// Tests/T_SafeTof_Tests
FUNCTION_BLOCK T_SafeTof_Tests EXTENDS TcUnit.FB_TestSuite
VAR
    // Test_OutputDelayedOff
    group_1 : T_SafeGroup;
    fb_1 : T_SafeTof(group := group_1) := (Parameters := (DelayTime := T#100MS));
    state_1 : INT := 10;
    waitTimer_1 : TON;
    // Test_UnconnectedInputIsRefused
    group_2 : T_SafeGroup;
    fb_2 : T_SafeTof(group := group_2);
END_VAR

Test_OutputDelayedOff();
Test_UnconnectedInputIsRefused();

METHOD PRIVATE Test_OutputDelayedOff
TcUnit.TEST(__POUNAME());
waitTimer_1();

CASE state_1 OF
    10:
        group_1(Run := TRUE);
        fb_1(TofIn1 := TRUE);
        AssertEquals_BOOL(Expected := TRUE, Actual := fb_1.TofOut, Message := 'output on immediately');
        // act
        fb_1(TofIn1 := FALSE);
        AssertEquals_BOOL(Expected := TRUE, Actual := fb_1.TofOut, Message := 'output held during the delay');
        AssertEquals_BYTE(Expected := TO_BYTE(E_SafeFbState.DelayOut), Actual := fb_1.State, Message := 'state DELAYOUT');
        state_1 := 20;
        waitTimer_1(IN := TRUE, PT := T#200MS);
    20:
        group_1(Run := TRUE);
        fb_1(TofIn1 := FALSE);

        IF NOT waitTimer_1.Q THEN
            RETURN;
        END_IF

        waitTimer_1(IN := FALSE);
        // assert
        AssertEquals_BOOL(Expected := FALSE, Actual := fb_1.TofOut, Message := 'output off after the delay');
        TEST_FINISHED_NAMED(__POUNAME());
        state_1 := 10;
END_CASE
END_METHOD

METHOD PRIVATE Test_UnconnectedInputIsRefused
TcUnit.TEST(__POUNAME());
// arrange / act: TofIn1 is unconnected, which the Safety Editor refuses
group_2(Run := TRUE);
fb_2();
group_2(Run := TRUE);
fb_2();
// assert
AssertEquals_BOOL(Expected := TRUE, Actual := fb_2.Error, Message := 'configuration error reported');
AssertEquals_BYTE(Expected := TO_BYTE(E_SafeFbState.Error), Actual := fb_2.State, Message := 'state ERROR');
AssertEquals_WORD(Expected := WORD#16#8000, Actual := fb_2.Diag, Message := 'diag bit 15 configuration refused');
AssertEquals_BOOL(Expected := FALSE, Actual := fb_2.TofOut, Message := 'TofOut stays at its safe value');
AssertEquals_BOOL(Expected := TRUE, Actual := group_2.FbErr, Message := 'the group sees an FB error');
// act: ErrAck 0 -> 1 -> 0 does not clear a configuration error
group_2(Run := TRUE, ErrAck := TRUE);
fb_2();
group_2(Run := TRUE, ErrAck := TRUE);
fb_2();
group_2(Run := TRUE, ErrAck := FALSE);
fb_2();
AssertEquals_BOOL(Expected := TRUE, Actual := fb_2.Error, Message := 'error not acknowledged');
AssertEquals_WORD(Expected := WORD#16#8000, Actual := fb_2.Diag, Message := 'diag bit 15 kept');
TEST_FINISHED_NAMED(__POUNAME());
END_METHOD

END_FUNCTION_BLOCK

// Tests/T_SafeEdm_Tests
FUNCTION_BLOCK T_SafeEdm_Tests EXTENDS TcUnit.FB_TestSuite
VAR
    // Test_SwitchOnTimeoutGivesError
    group_1 : T_SafeGroup;
    fb_1 : T_SafeEdm(group := group_1) := (Parameters := (SwitchOnTime := T#100MS));
    state_1 : INT := 10;
    waitTimer_1 : TON;
    // Test_NoErrorWhenFeedbackFollows
    group_2 : T_SafeGroup;
    fb_2 : T_SafeEdm(group := group_2) := (Parameters := (SwitchOnTime := T#100MS, SwitchOffTime := T#100MS));
    state_2 : INT := 10;
    waitTimer_2 : TON;
    // Test_UnconnectedMon2IsRefused
    group_3 : T_SafeGroup;
    fb_3 : T_SafeEdm(group := group_3);
END_VAR

Test_SwitchOnTimeoutGivesError();
Test_NoErrorWhenFeedbackFollows();
Test_UnconnectedMon2IsRefused();

METHOD PRIVATE Test_NoErrorWhenFeedbackFollows
TcUnit.TEST(__POUNAME());
waitTimer_2();

CASE state_2 OF
    10:
        state_2 := 20;
        waitTimer_2(IN := TRUE, PT := T#200MS);
    20:
        group_2(Run := TRUE);
        fb_2(Mon1 := TRUE, Mon2 := FALSE);

        IF NOT waitTimer_2.Q THEN
            RETURN;
        END_IF

        waitTimer_2(IN := FALSE);
        AssertEquals_BOOL(Expected := FALSE, Actual := fb_2.Error, Message := 'no error while feedback is correct');
        state_2 := 30;
        waitTimer_2(IN := TRUE, PT := T#200MS);
    30:
        // act: switch off, feedback follows immediately
        group_2(Run := TRUE);
        fb_2(Mon1 := FALSE, Mon2 := TRUE);

        IF NOT waitTimer_2.Q THEN
            RETURN;
        END_IF

        waitTimer_2(IN := FALSE);
        AssertEquals_BOOL(Expected := FALSE, Actual := fb_2.Error, Message := 'no error after switch-off with feedback');
        TEST_FINISHED_NAMED(__POUNAME());
        state_2 := 10;
END_CASE
END_METHOD

METHOD PRIVATE Test_SwitchOnTimeoutGivesError
TcUnit.TEST(__POUNAME());
waitTimer_1();

CASE state_1 OF
    10:
        state_1 := 20;
        waitTimer_1(IN := TRUE, PT := T#250MS);
    20:
        // act: Mon1 on, feedback never follows
        group_1(Run := TRUE, ErrAck := FALSE);
        fb_1(Mon1 := TRUE, Mon2 := TRUE);

        IF NOT waitTimer_1.Q THEN
            RETURN;
        END_IF

        waitTimer_1(IN := FALSE);
        // assert
        AssertEquals_BOOL(Expected := TRUE, Actual := fb_1.Error, Message := 'error when Mon2 does not drop in time');
        AssertEquals_WORD(Expected := WORD#2, Actual := fb_1.Diag, Message := 'diag bit 1 switch-on timer elapsed');
        // act: acknowledge (two cycles raised so the group_1 reaches RESET, then released)
        group_1(Run := TRUE, ErrAck := TRUE);
        fb_1(Mon1 := TRUE, Mon2 := TRUE);
        group_1(Run := TRUE, ErrAck := TRUE);
        fb_1(Mon1 := TRUE, Mon2 := TRUE);
        group_1(Run := TRUE, ErrAck := FALSE);
        fb_1(Mon1 := TRUE, Mon2 := FALSE);
        AssertEquals_BOOL(Expected := FALSE, Actual := fb_1.Error, Message := 'error cleared after acknowledgement');
        TEST_FINISHED_NAMED(__POUNAME());
        state_1 := 10;
END_CASE
END_METHOD

METHOD PRIVATE Test_UnconnectedMon2IsRefused
TcUnit.TEST(__POUNAME());
// arrange / act: Mon2 is unconnected, which the Safety Editor refuses
group_3(Run := TRUE);
fb_3(Mon1 := TRUE);
group_3(Run := TRUE);
fb_3(Mon1 := TRUE);
// assert
AssertEquals_BOOL(Expected := TRUE, Actual := fb_3.Error, Message := 'configuration error reported');
AssertEquals_BYTE(Expected := TO_BYTE(E_SafeFbState.Error), Actual := fb_3.State, Message := 'state ERROR');
AssertEquals_WORD(Expected := WORD#16#8000, Actual := fb_3.Diag, Message := 'diag bit 15 configuration refused');
AssertEquals_BOOL(Expected := TRUE, Actual := group_3.FbErr, Message := 'the group sees an FB error');
// act: ErrAck 0 -> 1 -> 0 does not clear a configuration error
group_3(Run := TRUE, ErrAck := TRUE);
fb_3(Mon1 := TRUE);
group_3(Run := TRUE, ErrAck := TRUE);
fb_3(Mon1 := TRUE);
group_3(Run := TRUE, ErrAck := FALSE);
fb_3(Mon1 := TRUE);
AssertEquals_BOOL(Expected := TRUE, Actual := fb_3.Error, Message := 'error not acknowledged');
AssertEquals_WORD(Expected := WORD#16#8000, Actual := fb_3.Diag, Message := 'diag bit 15 kept');
TEST_FINISHED_NAMED(__POUNAME());
END_METHOD

END_FUNCTION_BLOCK

// Tests/T_SafeEStop_Tests
FUNCTION_BLOCK T_SafeEStop_Tests EXTENDS TcUnit.FB_TestSuite
VAR
    // Test_OutputsOffWhenStopped
    group_1 : T_SafeGroup;
    fb_1 : T_SafeEStop(group := group_1);
    // Test_StartupRequiresRestartSequence
    group_2 : T_SafeGroup;
    fb_2 : T_SafeEStop(group := group_2);
    // Test_EStopRequestSwitchesOutputsOffAndBlocksRestart
    group_3 : T_SafeGroup;
    fb_3 : T_SafeEStop(group := group_3);
    // Test_MakeContactInputRequestsSafeStateOnOne
    group_4 : T_SafeGroup;
    fb_4 : T_SafeEStop(group := group_4) := (Parameters := (EStopIn1MakeContact := TRUE));
    // Test_EdmErrorAtRestartAndAcknowledge
    group_5 : T_SafeGroup;
    fb_5 : T_SafeEStop(group := group_5);
    // Test_RestartHeldBeforeEStopGivesEdmError
    group_6 : T_SafeGroup;
    fb_6 : T_SafeEStop(group := group_6);
    // Test_DelayedOutput
    group_7 : T_SafeGroup;
    fb_7 : T_SafeEStop(group := group_7) := (Parameters := (DelayTime := T#150MS));
    state_7 : INT := 10;
    waitTimer_7 : TON;
    // Test_DiscrepancyErrorNeedsSafeInputsBeforeAck
    group_8 : T_SafeGroup;
    fb_8 : T_SafeEStop(group := group_8) := (Parameters := (DiscrepancyTime1 := T#100MS));
    state_8 : INT := 10;
    waitTimer_8 : TON;
    // Test_ResetTimeOverSixtySecondsIsRefused
    group_9 : T_SafeGroup;
    fb_9 : T_SafeEStop(group := group_9) := (Parameters := (Edm2ResetTime := T#60010MS));
END_VAR

Test_OutputsOffWhenStopped();
Test_StartupRequiresRestartSequence();
Test_EStopRequestSwitchesOutputsOffAndBlocksRestart();
Test_MakeContactInputRequestsSafeStateOnOne();
Test_EdmErrorAtRestartAndAcknowledge();
Test_RestartHeldBeforeEStopGivesEdmError();
Test_DelayedOutput();
Test_DiscrepancyErrorNeedsSafeInputsBeforeAck();
Test_ResetTimeOverSixtySecondsIsRefused();

METHOD PRIVATE Test_DelayedOutput
TcUnit.TEST(__POUNAME());
waitTimer_7();

CASE state_7 OF
    10:
        // arrange: running
        group_7(Run := TRUE);
        fb_7(Restart := FALSE, EStopIn1 := TRUE);
        group_7(Run := TRUE);
        fb_7(Restart := TRUE, EStopIn1 := TRUE);
        group_7(Run := TRUE);
        fb_7(Restart := FALSE, EStopIn1 := TRUE);
        // act
        group_7(Run := TRUE);
        fb_7(Restart := FALSE, EStopIn1 := FALSE);
        // assert
        AssertEquals_BOOL(Expected := FALSE, Actual := fb_7.EStopOut, Message := 'EStopOut off immediately');
        AssertEquals_BOOL(Expected := TRUE, Actual := fb_7.EStopDelOut, Message := 'EStopDelOut still on');
        AssertEquals_BYTE(Expected := TO_BYTE(E_SafeFbState.DelayOut), Actual := fb_7.State, Message := 'state DELAYOUT');
        state_7 := 20;
        waitTimer_7(IN := TRUE, PT := T#300MS);
    20:
        group_7(Run := TRUE);
        fb_7(Restart := FALSE, EStopIn1 := FALSE);

        IF NOT waitTimer_7.Q THEN
            RETURN;
        END_IF

        waitTimer_7(IN := FALSE);
        // assert
        AssertEquals_BOOL(Expected := FALSE, Actual := fb_7.EStopDelOut, Message := 'EStopDelOut off after the delay');
        AssertEquals_BYTE(Expected := TO_BYTE(E_SafeFbState.Safe), Actual := fb_7.State, Message := 'state SAFE');
        TEST_FINISHED_NAMED(__POUNAME());
        state_7 := 10;
END_CASE
END_METHOD

METHOD PRIVATE Test_DiscrepancyErrorNeedsSafeInputsBeforeAck
TcUnit.TEST(__POUNAME());
waitTimer_8();

CASE state_8 OF
    10:
        // arrange: running
        group_8(Run := TRUE, ErrAck := FALSE);
        fb_8(Restart := FALSE, EStopIn1 := TRUE, EStopIn2 := TRUE);
        group_8(Run := TRUE, ErrAck := FALSE);
        fb_8(Restart := TRUE, EStopIn1 := TRUE, EStopIn2 := TRUE);
        group_8(Run := TRUE, ErrAck := FALSE);
        fb_8(Restart := FALSE, EStopIn1 := TRUE, EStopIn2 := TRUE);
        state_8 := 20;
        waitTimer_8(IN := TRUE, PT := T#250MS);
    20:
        // act: only one channel opens
        group_8(Run := TRUE, ErrAck := FALSE);
        fb_8(Restart := FALSE, EStopIn1 := FALSE, EStopIn2 := TRUE);

        IF NOT waitTimer_8.Q THEN
            RETURN;
        END_IF

        waitTimer_8(IN := FALSE);
        // assert
        AssertEquals_BOOL(Expected := TRUE, Actual := fb_8.Error, Message := 'discrepancy error');
        AssertEquals_WORD(Expected := WORD#16#0101, Actual := fb_8.Diag, Message := 'diag bits 0 and 8');
        // act: acknowledge while channel 2 is still closed
        group_8(Run := TRUE, ErrAck := TRUE);
        fb_8(Restart := FALSE, EStopIn1 := FALSE, EStopIn2 := TRUE);
        AssertEquals_BYTE(Expected := TO_BYTE(E_SafeFbState.Error), Actual := fb_8.State, Message := 'ack refused until both channels safe');
        group_8(Run := TRUE, ErrAck := TRUE);
        fb_8(Restart := FALSE, EStopIn1 := FALSE, EStopIn2 := FALSE);
        AssertEquals_BYTE(Expected := TO_BYTE(E_SafeFbState.Reset), Actual := fb_8.State, Message := 'RESET once both channels were safe');
        TEST_FINISHED_NAMED(__POUNAME());
        state_8 := 10;
END_CASE
END_METHOD

METHOD PRIVATE Test_EdmErrorAtRestartAndAcknowledge
TcUnit.TEST(__POUNAME());
// arrange: EDM1 connected but contactor not released
group_5(Run := TRUE, ErrAck := FALSE);
fb_5(Restart := FALSE, EDM1 := FALSE, EStopIn1 := TRUE);
// act: restart
group_5(Run := TRUE, ErrAck := FALSE);
fb_5(Restart := TRUE, EDM1 := FALSE, EStopIn1 := TRUE);
// assert
AssertEquals_BOOL(Expected := TRUE, Actual := fb_5.Error, Message := 'EDM error when feedback missing at restart');
AssertEquals_BYTE(Expected := TO_BYTE(E_SafeFbState.Error), Actual := fb_5.State, Message := 'state ERROR');
AssertEquals_WORD(Expected := WORD#16, Actual := fb_5.Diag, Message := 'diag bit 4 EDM1');
// act: the group_5 sees the error and leaves RUN; the FB error is held
group_5(Run := TRUE, ErrAck := FALSE);
fb_5(Restart := FALSE, EDM1 := FALSE, EStopIn1 := TRUE);
AssertEquals_BYTE(Expected := TO_BYTE(E_SafeGroupState.Error), Actual := group_5.State, Message := 'group ERROR');
AssertEquals_BYTE(Expected := TO_BYTE(E_SafeFbState.Error), Actual := fb_5.State, Message := 'error is held while the group is in ERROR');
// act: ErrAck 0 -> 1 (two cycles, the group_5 needs the second to reach RESET) -> 0
group_5(Run := TRUE, ErrAck := TRUE);
fb_5(Restart := FALSE, EDM1 := FALSE, EStopIn1 := TRUE);
AssertEquals_BYTE(Expected := TO_BYTE(E_SafeFbState.Reset), Actual := fb_5.State, Message := 'state RESET while ErrAck is 1');
AssertEquals_BOOL(Expected := FALSE, Actual := fb_5.Error, Message := 'Error output off in RESET');
group_5(Run := TRUE, ErrAck := TRUE);
fb_5(Restart := FALSE, EDM1 := FALSE, EStopIn1 := TRUE);
AssertEquals_BYTE(Expected := TO_BYTE(E_SafeGroupState.Reset), Actual := group_5.State, Message := 'group RESET');
group_5(Run := TRUE, ErrAck := FALSE);
fb_5(Restart := FALSE, EDM1 := FALSE, EStopIn1 := TRUE);
AssertEquals_BYTE(Expected := TO_BYTE(E_SafeGroupState.Run), Actual := group_5.State, Message := 'group RUN after ErrAck falling edge');
AssertEquals_BYTE(Expected := TO_BYTE(E_SafeFbState.Safe), Actual := fb_5.State, Message := 'state SAFE after ErrAck falling edge');
TEST_FINISHED_NAMED(__POUNAME());
END_METHOD

